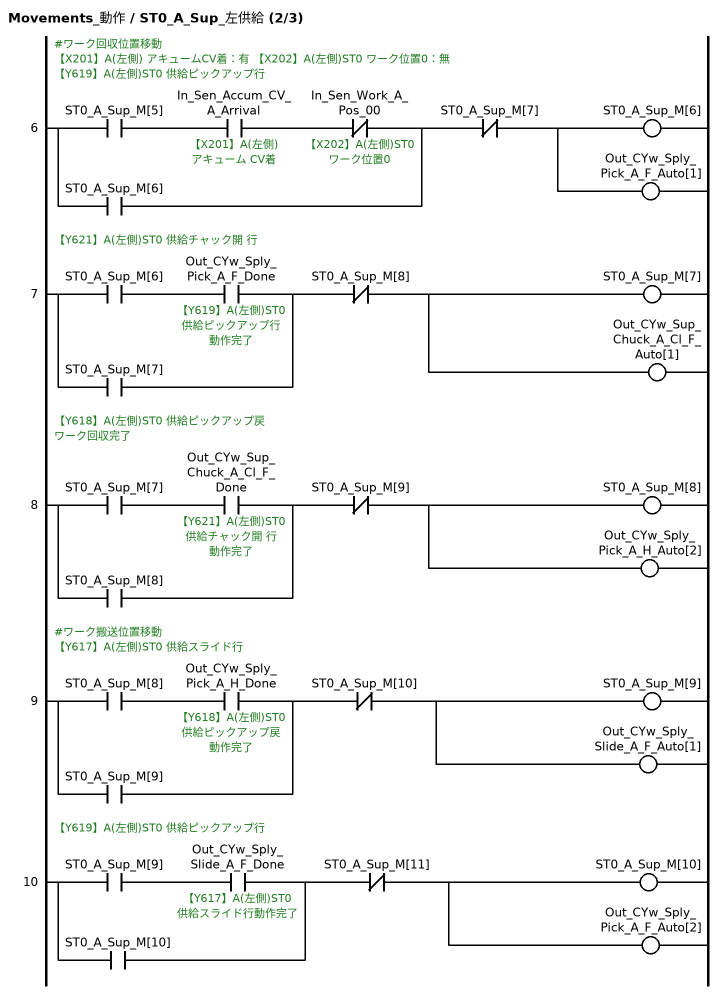
(* [picture p24: Movements_動作 / ST0_A_Sup_左供給, rungs 6-10] *)
(* Rung 6: #ワーク回収位置移動 / 【X201】A(左側) アキュームCV着：有 【X202】A(左側)ST0 ワーク位置0：無 / 【Y619】A(左側)ST0 供給ピックアップ行 *)
_p20 := ((ST0_A_Sup_M[5] AND In_Sen_Accum_CV_A_Arrival AND NOT In_Sen_Work_A_Pos_00) OR ST0_A_Sup_M[6]) AND NOT ST0_A_Sup_M[7];
ST0_A_Sup_M[6] := _p20;
Out_CYw_Sply_Pick_A_F_Auto[1] := _p20;
(* Rung 7: 【Y621】A(左側)ST0 供給チャック開 行 *)
_p21 := ((ST0_A_Sup_M[6] AND Out_CYw_Sply_Pick_A_F_Done) OR ST0_A_Sup_M[7]) AND NOT ST0_A_Sup_M[8];
ST0_A_Sup_M[7] := _p21;
Out_CYw_Sup_Chuck_A_Cl_F_Auto[1] := _p21;
(* Rung 8: 【Y618】A(左側)ST0 供給ピックアップ戻 / ワーク回収完了 *)
_p22 := ((ST0_A_Sup_M[7] AND Out_CYw_Sup_Chuck_A_Cl_F_Done) OR ST0_A_Sup_M[8]) AND NOT ST0_A_Sup_M[9];
ST0_A_Sup_M[8] := _p22;
Out_CYw_Sply_Pick_A_H_Auto[2] := _p22;
(* Rung 9: #ワーク搬送位置移動 / 【Y617】A(左側)ST0 供給スライド行 *)
_p23 := ((ST0_A_Sup_M[8] AND Out_CYw_Sply_Pick_A_H_Done) OR ST0_A_Sup_M[9]) AND NOT ST0_A_Sup_M[10];
ST0_A_Sup_M[9] := _p23;
Out_CYw_Sply_Slide_A_F_Auto[1] := _p23;
(* Rung 10: 【Y619】A(左側)ST0 供給ピックアップ行 *)
_p24 := ((ST0_A_Sup_M[9] AND Out_CYw_Sply_Slide_A_F_Done) OR ST0_A_Sup_M[10]) AND NOT ST0_A_Sup_M[11];
ST0_A_Sup_M[10] := _p24;
Out_CYw_Sply_Pick_A_F_Auto[2] := _p24;

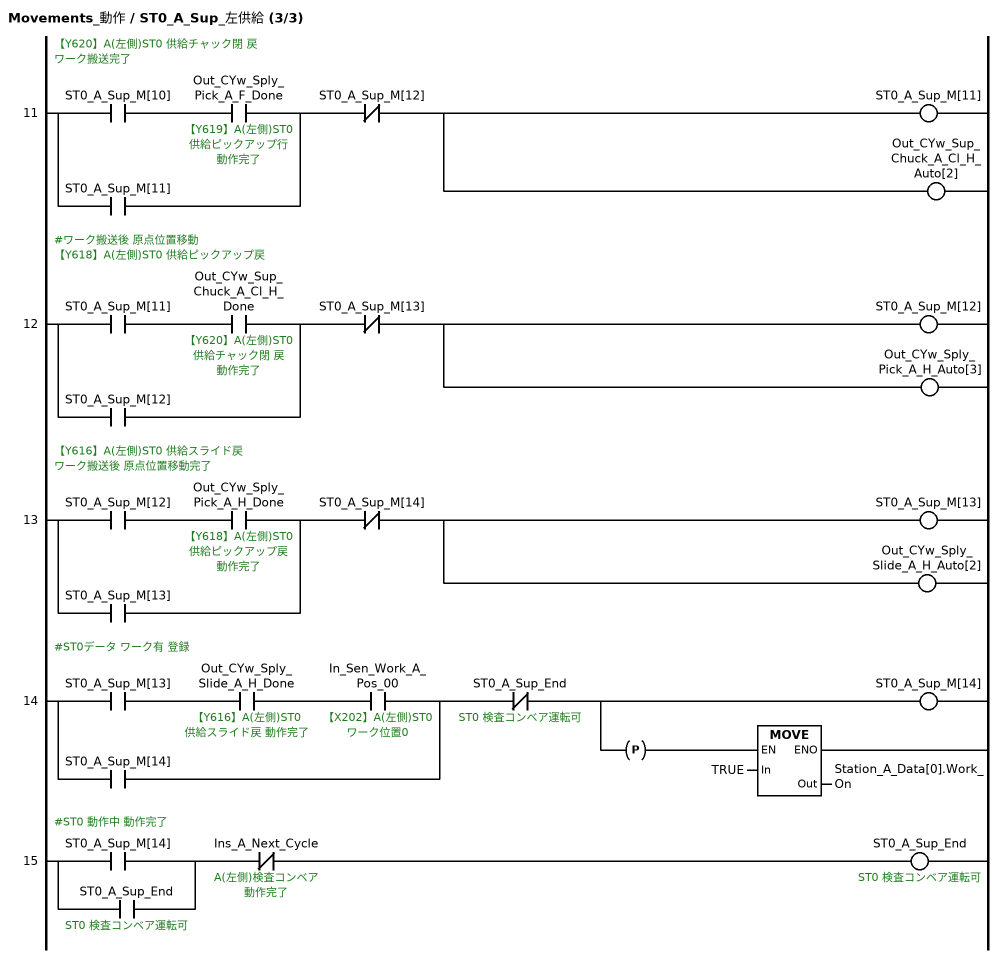
(* Rung 11: 【Y620】A(左側)ST0 供給チャック閉 戻 / ワーク搬送完了 *)
_p25 := ((ST0_A_Sup_M[10] AND Out_CYw_Sply_Pick_A_F_Done) OR ST0_A_Sup_M[11]) AND NOT ST0_A_Sup_M[12];
ST0_A_Sup_M[11] := _p25;
Out_CYw_Sup_Chuck_A_Cl_H_Auto[2] := _p25;
(* Rung 12: #ワーク搬送後 原点位置移動 / 【Y618】A(左側)ST0 供給ピックアップ戻 *)
_p26 := ((ST0_A_Sup_M[11] AND Out_CYw_Sup_Chuck_A_Cl_H_Done) OR ST0_A_Sup_M[12]) AND NOT ST0_A_Sup_M[13];
ST0_A_Sup_M[12] := _p26;
Out_CYw_Sply_Pick_A_H_Auto[3] := _p26;
(* Rung 13: 【Y616】A(左側)ST0 供給スライド戻 / ワーク搬送後 原点位置移動完了 *)
_p27 := ((ST0_A_Sup_M[12] AND Out_CYw_Sply_Pick_A_H_Done) OR ST0_A_Sup_M[13]) AND NOT ST0_A_Sup_M[14];
ST0_A_Sup_M[13] := _p27;
Out_CYw_Sply_Slide_A_H_Auto[2] := _p27;
(* Rung 14: #ST0データ ワーク有 登録 *)
_p28 := ((ST0_A_Sup_M[13] AND Out_CYw_Sply_Slide_A_H_Done AND In_Sen_Work_A_Pos_00) OR ST0_A_Sup_M[14]) AND NOT ST0_A_Sup_End;
ST0_A_Sup_M[14] := _p28;
_e29(CLK := _p28);
IF _e29.Q THEN Station_A_Data[0].Work_On := TRUE; END_IF;
(* Rung 15: #ST0 動作中 動作完了 *)
ST0_A_Sup_End := (ST0_A_Sup_M[14] OR ST0_A_Sup_End) AND NOT Ins_A_Next_Cycle;

(* Section ST1_A_Ca1_左Ca1検査: ladder, written here as Structured Text *)

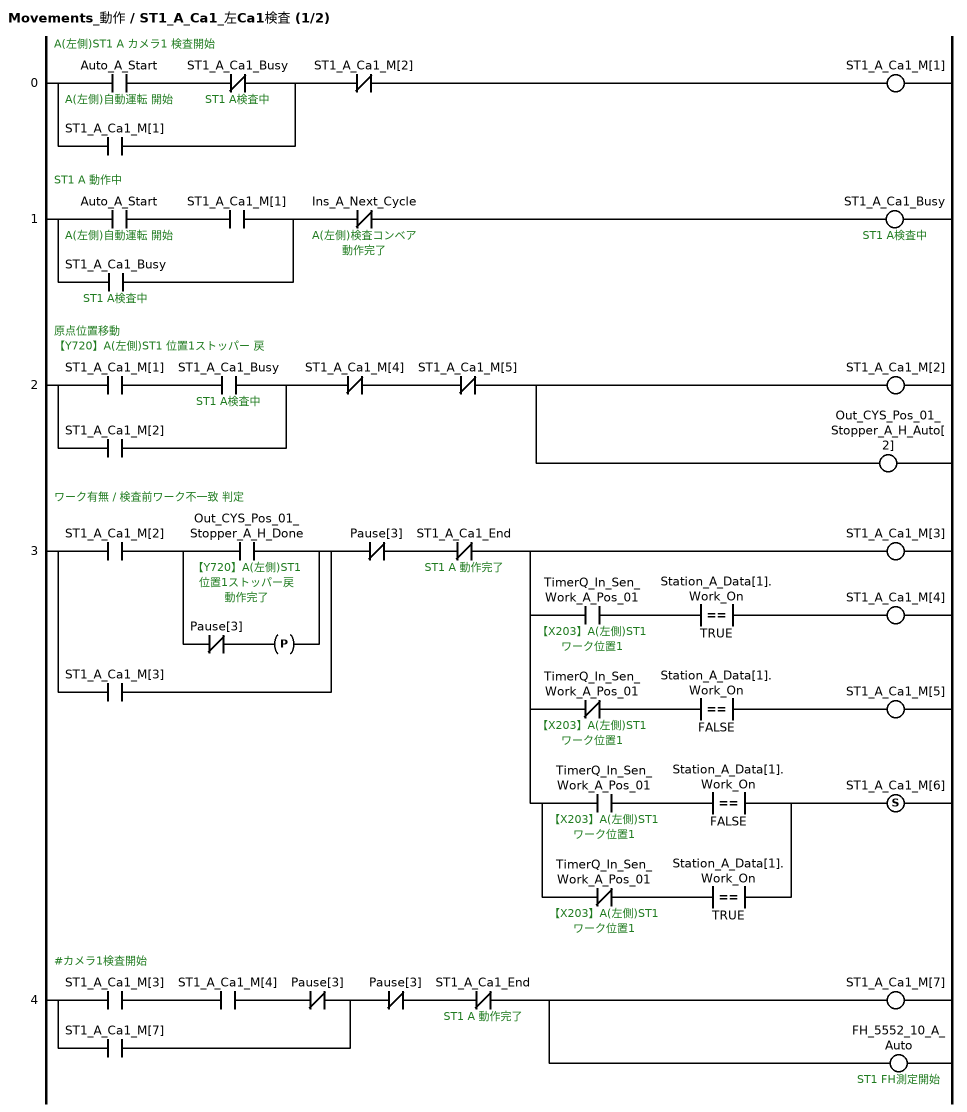
(* Rung 0: A(左側)ST1 A カメラ1 検査開始 *)
ST1_A_Ca1_M[1] := ((Auto_A_Start AND NOT ST1_A_Ca1_Busy) OR ST1_A_Ca1_M[1]) AND NOT ST1_A_Ca1_M[2];
(* Rung 1: ST1 A 動作中 *)
ST1_A_Ca1_Busy := ((Auto_A_Start AND ST1_A_Ca1_M[1]) OR ST1_A_Ca1_Busy) AND NOT Ins_A_Next_Cycle;
(* Rung 2: 原点位置移動 / 【Y720】A(左側)ST1 位置1ストッパー 戻 *)
_p30 := ((ST1_A_Ca1_M[1] AND ST1_A_Ca1_Busy) OR ST1_A_Ca1_M[2]) AND NOT ST1_A_Ca1_M[4] AND NOT ST1_A_Ca1_M[5];
ST1_A_Ca1_M[2] := _p30;
Out_CYS_Pos_01_Stopper_A_H_Auto[2] := _p30;
(* Rung 3: ワーク有無 / 検査前ワーク不一致 判定 *)
_e31(CLK := ST1_A_Ca1_M[2] AND NOT Pause[3]);
_p32 := ((ST1_A_Ca1_M[2] AND Out_CYS_Pos_01_Stopper_A_H_Done) OR _e31.Q OR ST1_A_Ca1_M[3]) AND NOT Pause[3] AND NOT ST1_A_Ca1_End;
ST1_A_Ca1_M[3] := _p32;
ST1_A_Ca1_M[4] := _p32 AND TimerQ_In_Sen_Work_A_Pos_01 AND (Station_A_Data[1].Work_On = TRUE);
ST1_A_Ca1_M[5] := _p32 AND NOT TimerQ_In_Sen_Work_A_Pos_01 AND (Station_A_Data[1].Work_On = FALSE);
IF _p32 AND ((TimerQ_In_Sen_Work_A_Pos_01 AND (Station_A_Data[1].Work_On = FALSE)) OR (NOT TimerQ_In_Sen_Work_A_Pos_01 AND (Station_A_Data[1].Work_On = TRUE))) THEN
    ST1_A_Ca1_M[6] := TRUE;
END_IF;
(* Rung 4: #カメラ1検査開始 *)
_p33 := ((ST1_A_Ca1_M[3] AND ST1_A_Ca1_M[4] AND NOT Pause[3]) OR ST1_A_Ca1_M[7]) AND NOT Pause[3] AND NOT ST1_A_Ca1_End;
ST1_A_Ca1_M[7] := _p33;
FH_5552_10_A_Auto := _p33;

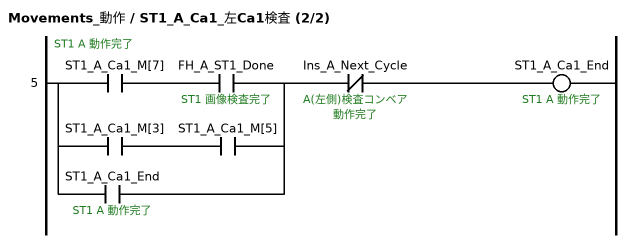
(* Rung 5: ST1 A 動作完了 *)
ST1_A_Ca1_End := ((ST1_A_Ca1_M[7] AND FH_A_ST1_Done) OR (ST1_A_Ca1_M[3] AND ST1_A_Ca1_M[5]) OR ST1_A_Ca1_End) AND NOT Ins_A_Next_Cycle;

(* Section ST2_A_Hgt_左高さ検査: ladder, written here as Structured Text *)

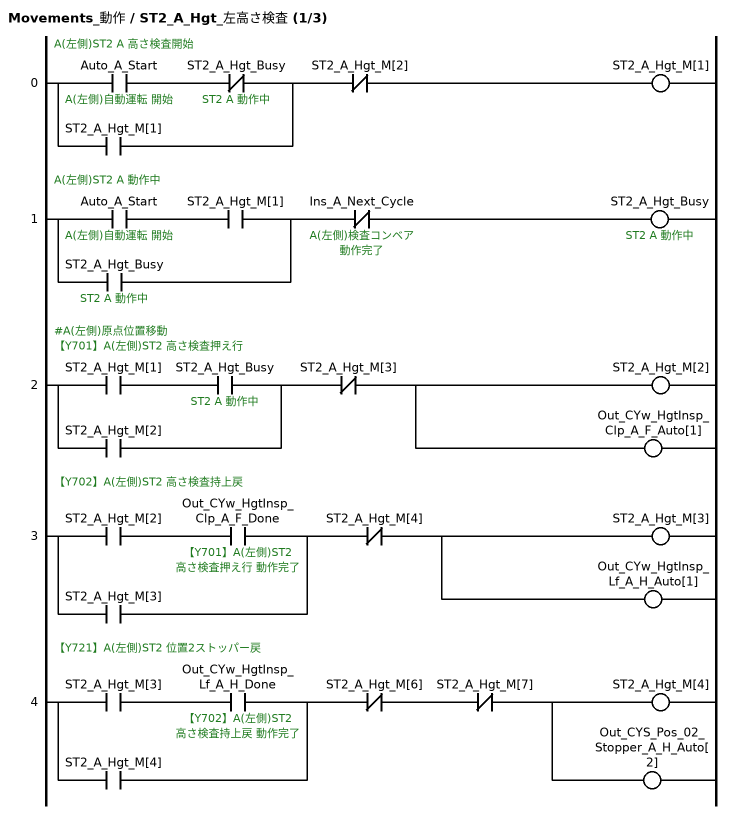
(* Rung 0: A(左側)ST2 A 高さ検査開始 *)
ST2_A_Hgt_M[1] := ((Auto_A_Start AND NOT ST2_A_Hgt_Busy) OR ST2_A_Hgt_M[1]) AND NOT ST2_A_Hgt_M[2];
(* Rung 1: A(左側)ST2 A 動作中 *)
ST2_A_Hgt_Busy := ((Auto_A_Start AND ST2_A_Hgt_M[1]) OR ST2_A_Hgt_Busy) AND NOT Ins_A_Next_Cycle;
(* Rung 2: #A(左側)原点位置移動 / 【Y701】A(左側)ST2 高さ検査押え行 *)
_p34 := ((ST2_A_Hgt_M[1] AND ST2_A_Hgt_Busy) OR ST2_A_Hgt_M[2]) AND NOT ST2_A_Hgt_M[3];
ST2_A_Hgt_M[2] := _p34;
Out_CYw_HgtInsp_Clp_A_F_Auto[1] := _p34;
(* Rung 3: 【Y702】A(左側)ST2 高さ検査持上戻 *)
_p35 := ((ST2_A_Hgt_M[2] AND Out_CYw_HgtInsp_Clp_A_F_Done) OR ST2_A_Hgt_M[3]) AND NOT ST2_A_Hgt_M[4];
ST2_A_Hgt_M[3] := _p35;
Out_CYw_HgtInsp_Lf_A_H_Auto[1] := _p35;
(* Rung 4: 【Y721】A(左側)ST2 位置2ストッパー戻 *)
_p36 := ((ST2_A_Hgt_M[3] AND Out_CYw_HgtInsp_Lf_A_H_Done) OR ST2_A_Hgt_M[4]) AND NOT ST2_A_Hgt_M[6] AND NOT ST2_A_Hgt_M[7];
ST2_A_Hgt_M[4] := _p36;
Out_CYS_Pos_02_Stopper_A_H_Auto[2] := _p36;

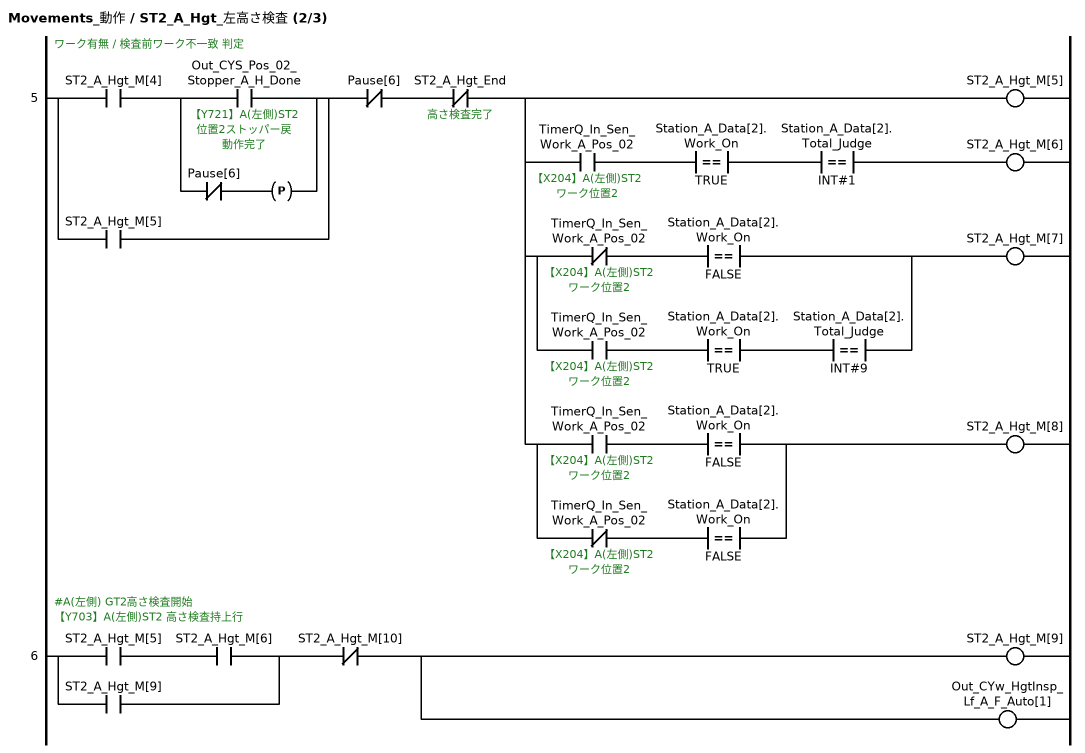
(* Rung 5: ワーク有無 / 検査前ワーク不一致 判定 *)
_e37(CLK := ST2_A_Hgt_M[4] AND NOT Pause[6]);
_p38 := ((ST2_A_Hgt_M[4] AND Out_CYS_Pos_02_Stopper_A_H_Done) OR _e37.Q OR ST2_A_Hgt_M[5]) AND NOT Pause[6] AND NOT ST2_A_Hgt_End;
ST2_A_Hgt_M[5] := _p38;
ST2_A_Hgt_M[6] := _p38 AND TimerQ_In_Sen_Work_A_Pos_02 AND (Station_A_Data[2].Work_On = TRUE) AND (Station_A_Data[2].Total_Judge = INT#1);
ST2_A_Hgt_M[7] := _p38 AND ((NOT TimerQ_In_Sen_Work_A_Pos_02 AND (Station_A_Data[2].Work_On = FALSE)) OR (TimerQ_In_Sen_Work_A_Pos_02 AND (Station_A_Data[2].Work_On = TRUE) AND (Station_A_Data[2].Total_Judge = INT#9)));
ST2_A_Hgt_M[8] := _p38 AND ((TimerQ_In_Sen_Work_A_Pos_02 AND (Station_A_Data[2].Work_On = FALSE)) OR (NOT TimerQ_In_Sen_Work_A_Pos_02 AND (Station_A_Data[2].Work_On = FALSE)));
(* Rung 6: #A(左側) GT2高さ検査開始 / 【Y703】A(左側)ST2 高さ検査持上行 *)
_p39 := ((ST2_A_Hgt_M[5] AND ST2_A_Hgt_M[6]) OR ST2_A_Hgt_M[9]) AND NOT ST2_A_Hgt_M[10];
ST2_A_Hgt_M[9] := _p39;
Out_CYw_HgtInsp_Lf_A_F_Auto[1] := _p39;

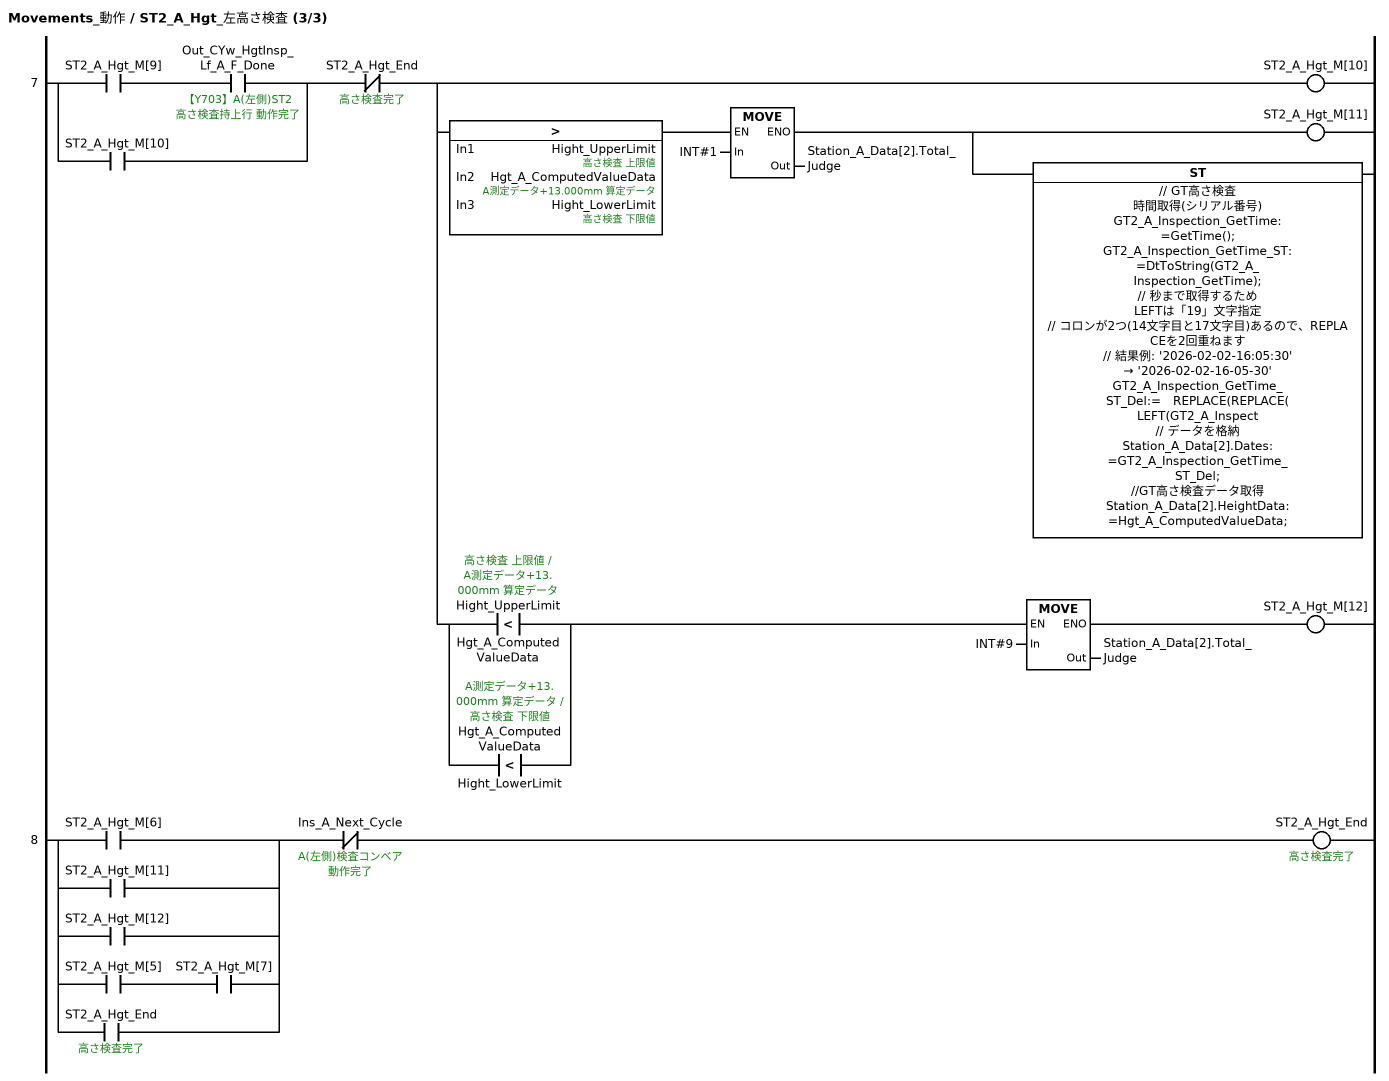
(* Rung 7 *)
_p40 := ((ST2_A_Hgt_M[9] AND Out_CYw_HgtInsp_Lf_A_F_Done) OR ST2_A_Hgt_M[10]) AND NOT ST2_A_Hgt_End;
ST2_A_Hgt_M[10] := _p40;
IF _p40 AND GT(Hight_UpperLimit, Hgt_A_ComputedValueData, Hight_LowerLimit) THEN
    Station_A_Data[2].Total_Judge := INT#1;
END_IF;
_p41 := _p40 AND GT(Hight_UpperLimit, Hgt_A_ComputedValueData, Hight_LowerLimit);
ST2_A_Hgt_M[11] := _p41;
IF _p41 THEN
    // GT高さ検査 時間取得(シリアル番号)
    GT2_A_Inspection_GetTime:=GetTime();
    GT2_A_Inspection_GetTime_ST:=DtToString(GT2_A_Inspection_GetTime);
    // 秒まで取得するため LEFTは「19」文字指定
    // コロンが2つ(14文字目と17文字目)あるので、REPLACEを2回重ねます
    // 結果例: '2026-02-02-16:05:30' → '2026-02-02-16-05-30'
    GT2_A_Inspection_GetTime_ST_Del:=   REPLACE(REPLACE(LEFT(GT2_A_Inspection_GetTime_ST, UINT#19), STRING#'-', UINT#1, UINT#17), STRING#'-', UINT#1, UINT#14);
    // データを格納
    Station_A_Data[2].Dates:=GT2_A_Inspection_GetTime_ST_Del;
    //GT高さ検査データ取得
    Station_A_Data[2].HeightData:=Hgt_A_ComputedValueData;
END_IF;
IF _p40 AND ((Hight_UpperLimit < Hgt_A_ComputedValueData) OR (Hgt_A_ComputedValueData < Hight_LowerLimit)) THEN
    Station_A_Data[2].Total_Judge := INT#9;
END_IF;
ST2_A_Hgt_M[12] := _p40 AND ((Hight_UpperLimit < Hgt_A_ComputedValueData) OR (Hgt_A_ComputedValueData < Hight_LowerLimit));
(* Rung 8 *)
ST2_A_Hgt_End := (ST2_A_Hgt_M[6] OR ST2_A_Hgt_M[11] OR ST2_A_Hgt_M[12] OR (ST2_A_Hgt_M[5] AND ST2_A_Hgt_M[7]) OR ST2_A_Hgt_End) AND NOT Ins_A_Next_Cycle;

(* Section ST3_A_Dis1_左NG1排出: ladder, written here as Structured Text *)

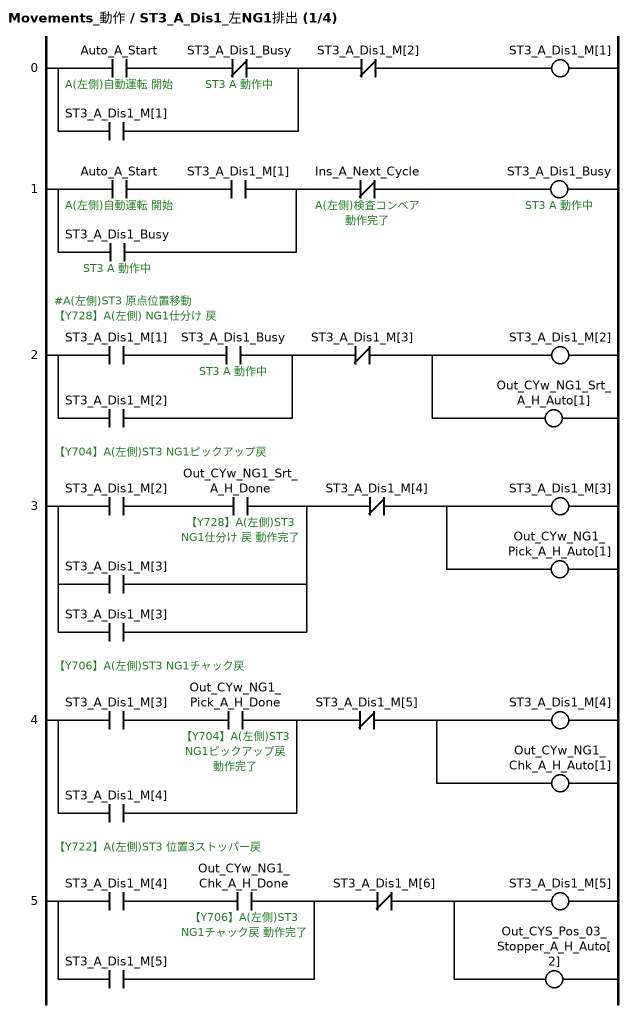
(* Rung 0 *)
ST3_A_Dis1_M[1] := ((Auto_A_Start AND NOT ST3_A_Dis1_Busy) OR ST3_A_Dis1_M[1]) AND NOT ST3_A_Dis1_M[2];
(* Rung 1 *)
ST3_A_Dis1_Busy := ((Auto_A_Start AND ST3_A_Dis1_M[1]) OR ST3_A_Dis1_Busy) AND NOT Ins_A_Next_Cycle;
(* Rung 2: #A(左側)ST3 原点位置移動 / 【Y728】A(左側) NG1仕分け 戻 *)
_p42 := ((ST3_A_Dis1_M[1] AND ST3_A_Dis1_Busy) OR ST3_A_Dis1_M[2]) AND NOT ST3_A_Dis1_M[3];
ST3_A_Dis1_M[2] := _p42;
Out_CYw_NG1_Srt_A_H_Auto[1] := _p42;
(* Rung 3: 【Y704】A(左側)ST3 NG1ピックアップ戻 *)
_p43 := ((ST3_A_Dis1_M[2] AND Out_CYw_NG1_Srt_A_H_Done) OR ST3_A_Dis1_M[3] OR ST3_A_Dis1_M[3]) AND NOT ST3_A_Dis1_M[4];
ST3_A_Dis1_M[3] := _p43;
Out_CYw_NG1_Pick_A_H_Auto[1] := _p43;
(* Rung 4: 【Y706】A(左側)ST3 NG1チャック戻 *)
_p44 := ((ST3_A_Dis1_M[3] AND Out_CYw_NG1_Pick_A_H_Done) OR ST3_A_Dis1_M[4]) AND NOT ST3_A_Dis1_M[5];
ST3_A_Dis1_M[4] := _p44;
Out_CYw_NG1_Chk_A_H_Auto[1] := _p44;
(* Rung 5: 【Y722】A(左側)ST3 位置3ストッパー戻 *)
_p45 := ((ST3_A_Dis1_M[4] AND Out_CYw_NG1_Chk_A_H_Done) OR ST3_A_Dis1_M[5]) AND NOT ST3_A_Dis1_M[6];
ST3_A_Dis1_M[5] := _p45;
Out_CYS_Pos_03_Stopper_A_H_Auto[2] := _p45;

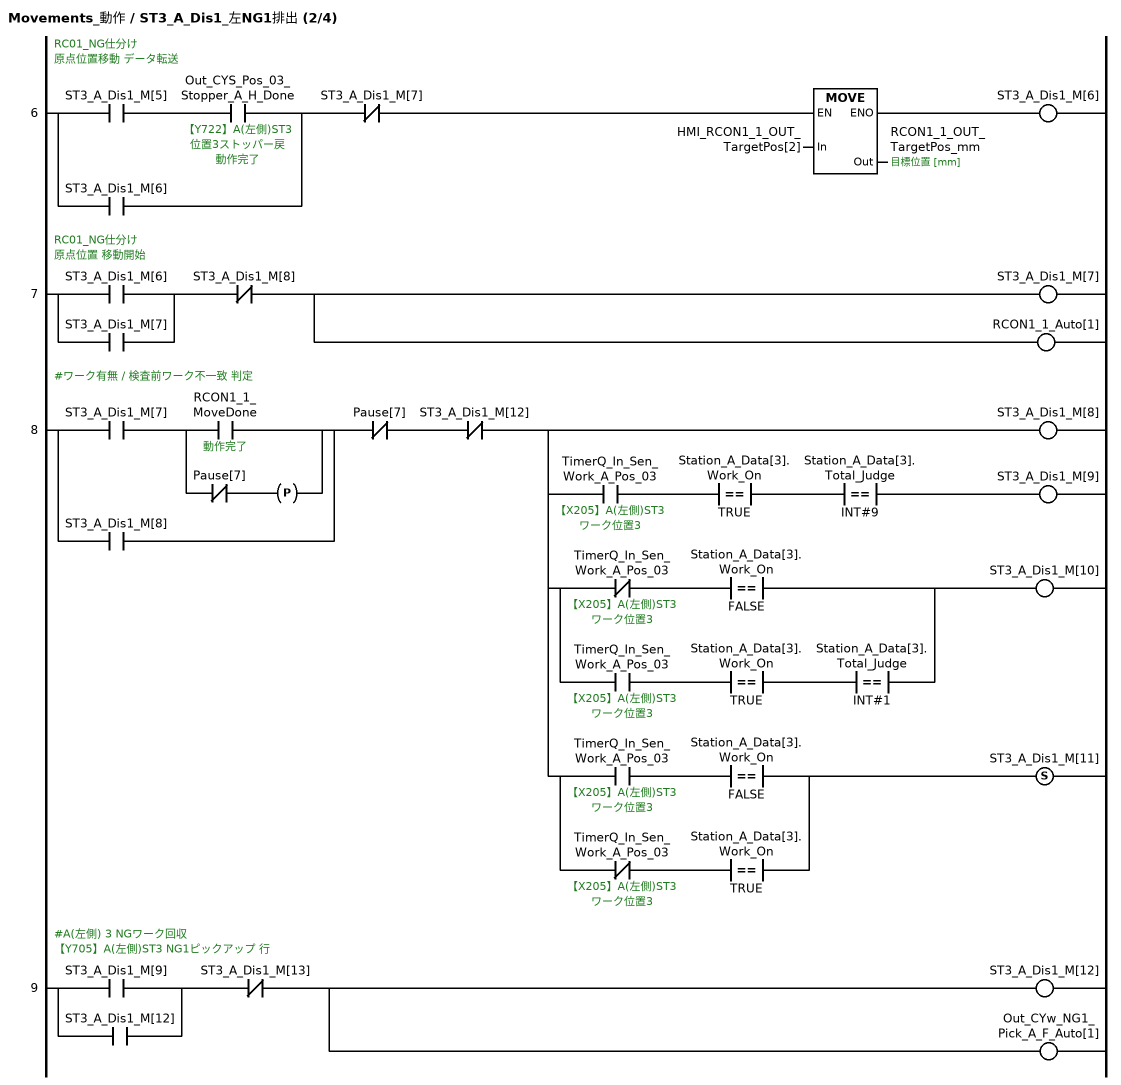
(* Rung 6: RC01_NG仕分け / 原点位置移動 データ転送 *)
IF ((ST3_A_Dis1_M[5] AND Out_CYS_Pos_03_Stopper_A_H_Done) OR ST3_A_Dis1_M[6]) AND NOT ST3_A_Dis1_M[7] THEN
    RCON1_1_OUT_TargetPos_mm := HMI_RCON1_1_OUT_TargetPos[2];
END_IF;
ST3_A_Dis1_M[6] := ((ST3_A_Dis1_M[5] AND Out_CYS_Pos_03_Stopper_A_H_Done) OR ST3_A_Dis1_M[6]) AND NOT ST3_A_Dis1_M[7];
(* Rung 7: RC01_NG仕分け / 原点位置 移動開始 *)
_p46 := (ST3_A_Dis1_M[6] OR ST3_A_Dis1_M[7]) AND NOT ST3_A_Dis1_M[8];
ST3_A_Dis1_M[7] := _p46;
RCON1_1_Auto[1] := _p46;
(* Rung 8: #ワーク有無 / 検査前ワーク不一致 判定 *)
_e47(CLK := ST3_A_Dis1_M[7] AND NOT Pause[7]);
_p48 := ((ST3_A_Dis1_M[7] AND RCON1_1_MoveDone) OR _e47.Q OR ST3_A_Dis1_M[8]) AND NOT Pause[7] AND NOT ST3_A_Dis1_M[12];
ST3_A_Dis1_M[8] := _p48;
ST3_A_Dis1_M[9] := _p48 AND TimerQ_In_Sen_Work_A_Pos_03 AND (Station_A_Data[3].Work_On = TRUE) AND (Station_A_Data[3].Total_Judge = INT#9);
ST3_A_Dis1_M[10] := _p48 AND ((NOT TimerQ_In_Sen_Work_A_Pos_03 AND (Station_A_Data[3].Work_On = FALSE)) OR (TimerQ_In_Sen_Work_A_Pos_03 AND (Station_A_Data[3].Work_On = TRUE) AND (Station_A_Data[3].Total_Judge = INT#1)));
IF _p48 AND ((TimerQ_In_Sen_Work_A_Pos_03 AND (Station_A_Data[3].Work_On = FALSE)) OR (NOT TimerQ_In_Sen_Work_A_Pos_03 AND (Station_A_Data[3].Work_On = TRUE))) THEN
    ST3_A_Dis1_M[11] := TRUE;
END_IF;
(* Rung 9: #A(左側) 3 NGワーク回収 / 【Y705】A(左側)ST3 NG1ピックアップ 行 *)
_p49 := (ST3_A_Dis1_M[9] OR ST3_A_Dis1_M[12]) AND NOT ST3_A_Dis1_M[13];
ST3_A_Dis1_M[12] := _p49;
Out_CYw_NG1_Pick_A_F_Auto[1] := _p49;

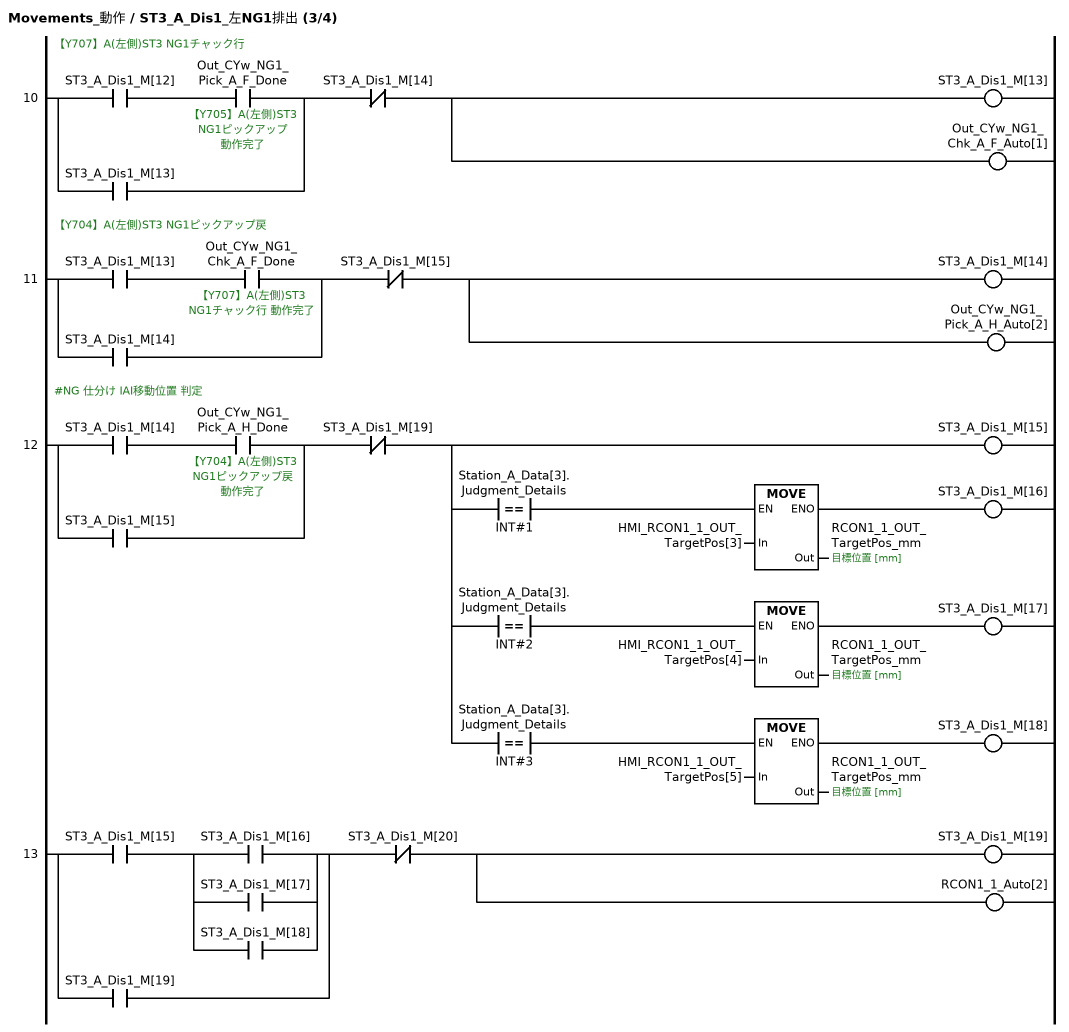
(* Rung 10: 【Y707】A(左側)ST3 NG1チャック行 *)
_p50 := ((ST3_A_Dis1_M[12] AND Out_CYw_NG1_Pick_A_F_Done) OR ST3_A_Dis1_M[13]) AND NOT ST3_A_Dis1_M[14];
ST3_A_Dis1_M[13] := _p50;
Out_CYw_NG1_Chk_A_F_Auto[1] := _p50;
(* Rung 11: 【Y704】A(左側)ST3 NG1ピックアップ戻 *)
_p51 := ((ST3_A_Dis1_M[13] AND Out_CYw_NG1_Chk_A_F_Done) OR ST3_A_Dis1_M[14]) AND NOT ST3_A_Dis1_M[15];
ST3_A_Dis1_M[14] := _p51;
Out_CYw_NG1_Pick_A_H_Auto[2] := _p51;
(* Rung 12: #NG 仕分け IAI移動位置 判定 *)
_p52 := ((ST3_A_Dis1_M[14] AND Out_CYw_NG1_Pick_A_H_Done) OR ST3_A_Dis1_M[15]) AND NOT ST3_A_Dis1_M[19];
ST3_A_Dis1_M[15] := _p52;
IF _p52 AND (Station_A_Data[3].Judgment_Details = INT#1) THEN
    RCON1_1_OUT_TargetPos_mm := HMI_RCON1_1_OUT_TargetPos[3];
END_IF;
ST3_A_Dis1_M[16] := _p52 AND (Station_A_Data[3].Judgment_Details = INT#1);
IF _p52 AND (Station_A_Data[3].Judgment_Details = INT#2) THEN
    RCON1_1_OUT_TargetPos_mm := HMI_RCON1_1_OUT_TargetPos[4];
END_IF;
ST3_A_Dis1_M[17] := _p52 AND (Station_A_Data[3].Judgment_Details = INT#2);
IF _p52 AND (Station_A_Data[3].Judgment_Details = INT#3) THEN
    RCON1_1_OUT_TargetPos_mm := HMI_RCON1_1_OUT_TargetPos[5];
END_IF;
ST3_A_Dis1_M[18] := _p52 AND (Station_A_Data[3].Judgment_Details = INT#3);
(* Rung 13 *)
_p53 := ((ST3_A_Dis1_M[15] AND (ST3_A_Dis1_M[16] OR ST3_A_Dis1_M[17] OR ST3_A_Dis1_M[18])) OR ST3_A_Dis1_M[19]) AND NOT ST3_A_Dis1_M[20];
ST3_A_Dis1_M[19] := _p53;
RCON1_1_Auto[2] := _p53;

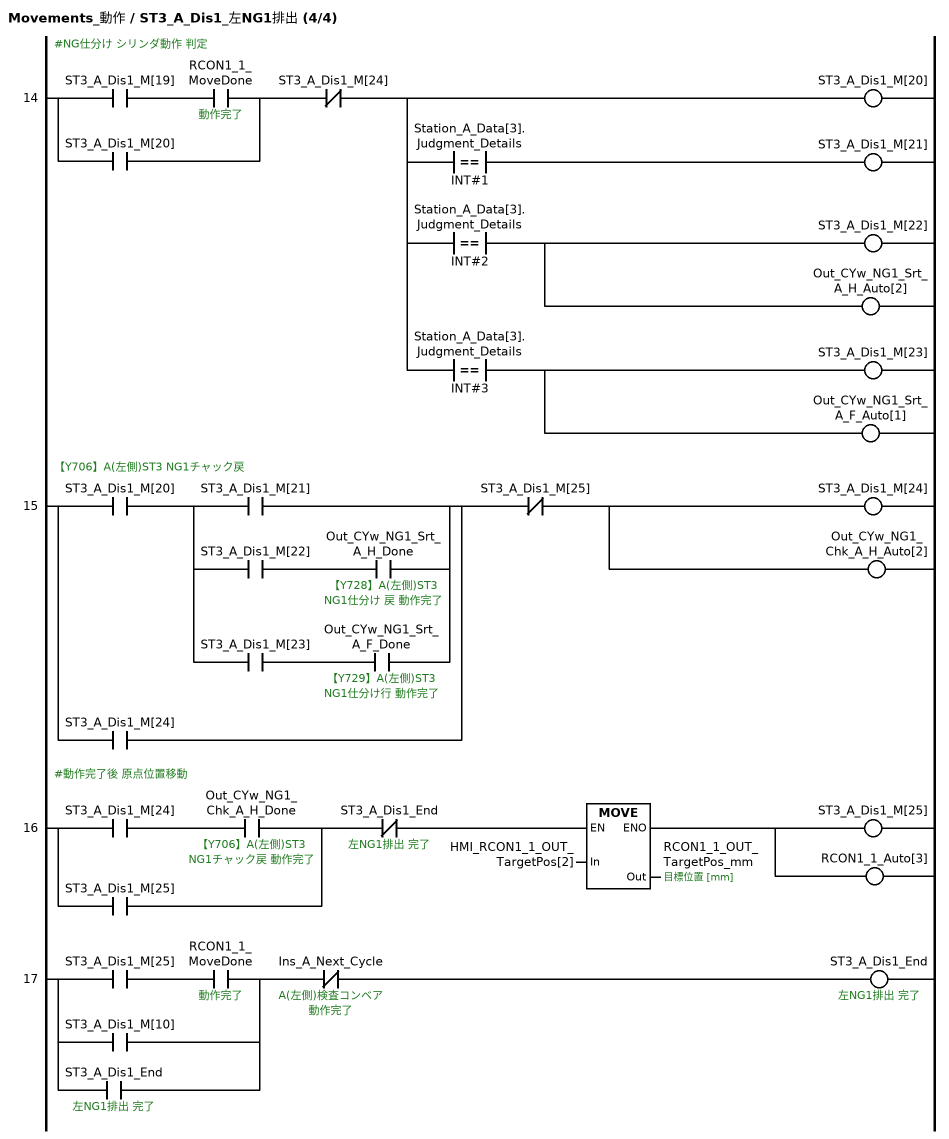
(* Rung 14: #NG仕分け シリンダ動作 判定 *)
_p54 := ((ST3_A_Dis1_M[19] AND RCON1_1_MoveDone) OR ST3_A_Dis1_M[20]) AND NOT ST3_A_Dis1_M[24];
ST3_A_Dis1_M[20] := _p54;
ST3_A_Dis1_M[21] := _p54 AND (Station_A_Data[3].Judgment_Details = INT#1);
_p55 := _p54 AND (Station_A_Data[3].Judgment_Details = INT#2);
ST3_A_Dis1_M[22] := _p55;
Out_CYw_NG1_Srt_A_H_Auto[2] := _p55;
_p56 := _p54 AND (Station_A_Data[3].Judgment_Details = INT#3);
ST3_A_Dis1_M[23] := _p56;
Out_CYw_NG1_Srt_A_F_Auto[1] := _p56;
(* Rung 15: 【Y706】A(左側)ST3 NG1チャック戻 *)
_p57 := ((ST3_A_Dis1_M[20] AND (ST3_A_Dis1_M[21] OR (ST3_A_Dis1_M[22] AND Out_CYw_NG1_Srt_A_H_Done) OR (ST3_A_Dis1_M[23] AND Out_CYw_NG1_Srt_A_F_Done))) OR ST3_A_Dis1_M[24]) AND NOT ST3_A_Dis1_M[25];
ST3_A_Dis1_M[24] := _p57;
Out_CYw_NG1_Chk_A_H_Auto[2] := _p57;
(* Rung 16: #動作完了後 原点位置移動 *)
IF ((ST3_A_Dis1_M[24] AND Out_CYw_NG1_Chk_A_H_Done) OR ST3_A_Dis1_M[25]) AND NOT ST3_A_Dis1_End THEN
    RCON1_1_OUT_TargetPos_mm := HMI_RCON1_1_OUT_TargetPos[2];
END_IF;
_p58 := ((ST3_A_Dis1_M[24] AND Out_CYw_NG1_Chk_A_H_Done) OR ST3_A_Dis1_M[25]) AND NOT ST3_A_Dis1_End;
ST3_A_Dis1_M[25] := _p58;
RCON1_1_Auto[3] := _p58;
(* Rung 17 *)
ST3_A_Dis1_End := ((ST3_A_Dis1_M[25] AND RCON1_1_MoveDone) OR ST3_A_Dis1_M[10] OR ST3_A_Dis1_End) AND NOT Ins_A_Next_Cycle;

(* Section ST4_A_Rev1_左反転1: ladder, written here as Structured Text *)

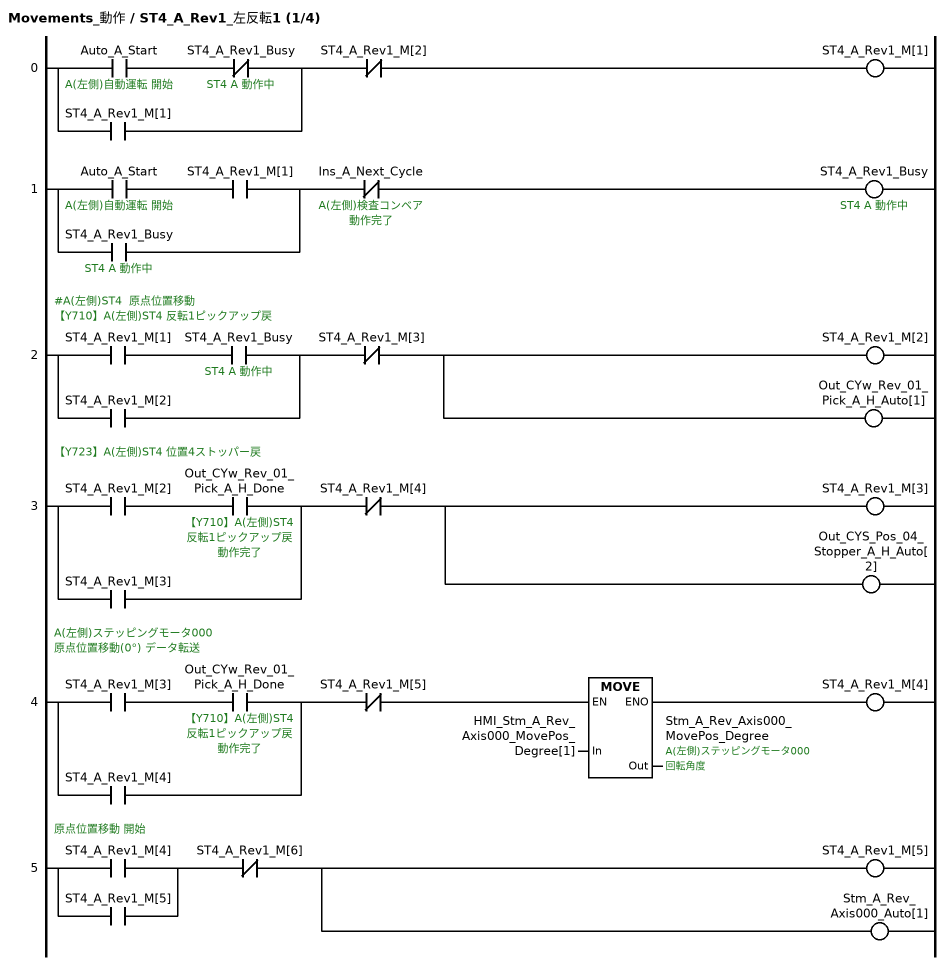
(* Rung 0 *)
ST4_A_Rev1_M[1] := ((Auto_A_Start AND NOT ST4_A_Rev1_Busy) OR ST4_A_Rev1_M[1]) AND NOT ST4_A_Rev1_M[2];
(* Rung 1 *)
ST4_A_Rev1_Busy := ((Auto_A_Start AND ST4_A_Rev1_M[1]) OR ST4_A_Rev1_Busy) AND NOT Ins_A_Next_Cycle;
(* Rung 2: #A(左側)ST4  原点位置移動 / 【Y710】A(左側)ST4 反転1ピックアップ戻 *)
_p59 := ((ST4_A_Rev1_M[1] AND ST4_A_Rev1_Busy) OR ST4_A_Rev1_M[2]) AND NOT ST4_A_Rev1_M[3];
ST4_A_Rev1_M[2] := _p59;
Out_CYw_Rev_01_Pick_A_H_Auto[1] := _p59;
(* Rung 3: 【Y723】A(左側)ST4 位置4ストッパー戻 *)
_p60 := ((ST4_A_Rev1_M[2] AND Out_CYw_Rev_01_Pick_A_H_Done) OR ST4_A_Rev1_M[3]) AND NOT ST4_A_Rev1_M[4];
ST4_A_Rev1_M[3] := _p60;
Out_CYS_Pos_04_Stopper_A_H_Auto[2] := _p60;
(* Rung 4: A(左側)ステッピングモータ000 / 原点位置移動(0°) データ転送 *)
IF ((ST4_A_Rev1_M[3] AND Out_CYw_Rev_01_Pick_A_H_Done) OR ST4_A_Rev1_M[4]) AND NOT ST4_A_Rev1_M[5] THEN
    Stm_A_Rev_Axis000_MovePos_Degree := HMI_Stm_A_Rev_Axis000_MovePos_Degree[1];
END_IF;
ST4_A_Rev1_M[4] := ((ST4_A_Rev1_M[3] AND Out_CYw_Rev_01_Pick_A_H_Done) OR ST4_A_Rev1_M[4]) AND NOT ST4_A_Rev1_M[5];
(* Rung 5: 原点位置移動 開始 *)
_p61 := (ST4_A_Rev1_M[4] OR ST4_A_Rev1_M[5]) AND NOT ST4_A_Rev1_M[6];
ST4_A_Rev1_M[5] := _p61;
Stm_A_Rev_Axis000_Auto[1] := _p61;

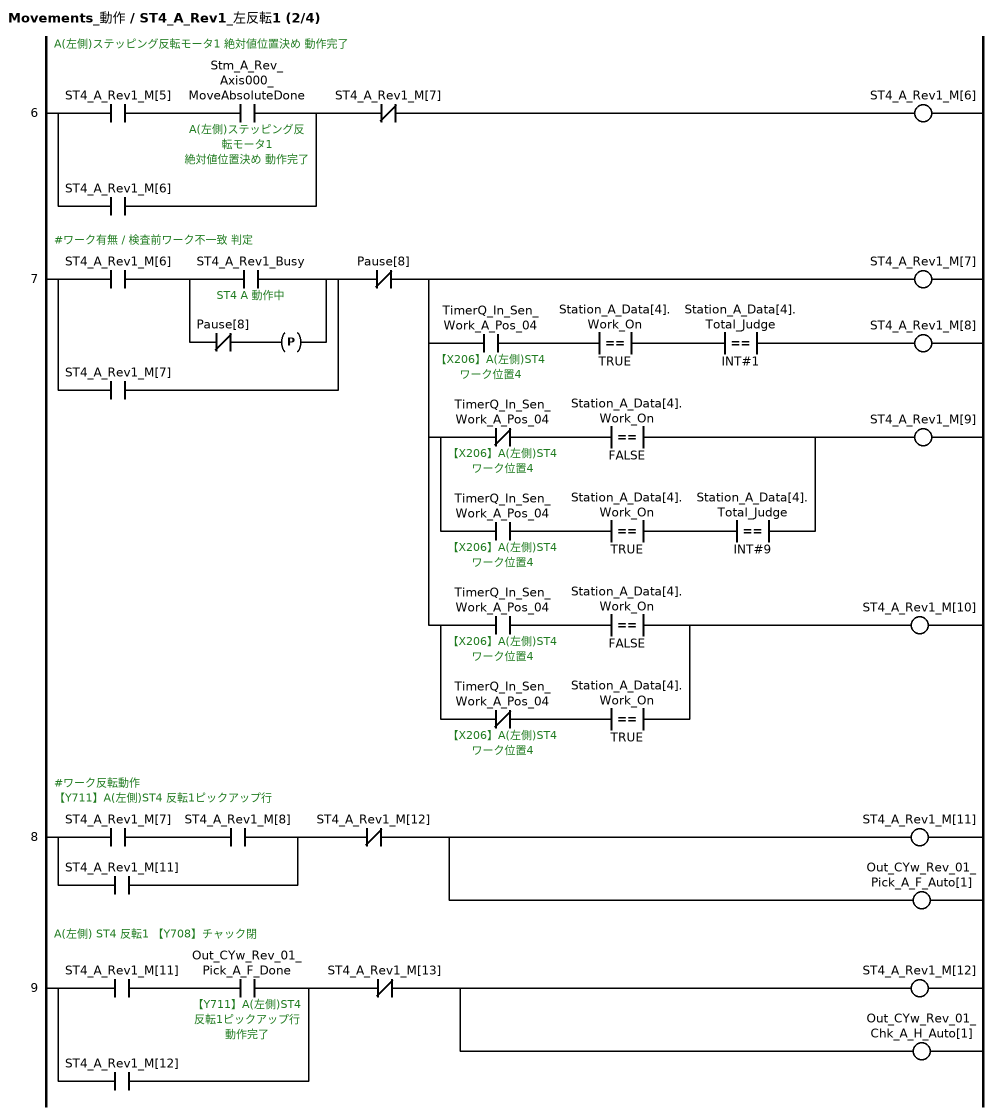
(* Rung 6: A(左側)ステッピング反転モータ1 絶対値位置決め 動作完了 *)
ST4_A_Rev1_M[6] := ((ST4_A_Rev1_M[5] AND Stm_A_Rev_Axis000_MoveAbsoluteDone) OR ST4_A_Rev1_M[6]) AND NOT ST4_A_Rev1_M[7];
(* Rung 7: #ワーク有無 / 検査前ワーク不一致 判定 *)
_e62(CLK := ST4_A_Rev1_M[6] AND NOT Pause[8]);
_p63 := ((ST4_A_Rev1_M[6] AND ST4_A_Rev1_Busy) OR _e62.Q OR ST4_A_Rev1_M[7]) AND NOT Pause[8];
ST4_A_Rev1_M[7] := _p63;
ST4_A_Rev1_M[8] := _p63 AND TimerQ_In_Sen_Work_A_Pos_04 AND (Station_A_Data[4].Work_On = TRUE) AND (Station_A_Data[4].Total_Judge = INT#1);
ST4_A_Rev1_M[9] := _p63 AND ((NOT TimerQ_In_Sen_Work_A_Pos_04 AND (Station_A_Data[4].Work_On = FALSE)) OR (TimerQ_In_Sen_Work_A_Pos_04 AND (Station_A_Data[4].Work_On = TRUE) AND (Station_A_Data[4].Total_Judge = INT#9)));
ST4_A_Rev1_M[10] := _p63 AND ((TimerQ_In_Sen_Work_A_Pos_04 AND (Station_A_Data[4].Work_On = FALSE)) OR (NOT TimerQ_In_Sen_Work_A_Pos_04 AND (Station_A_Data[4].Work_On = TRUE)));
(* Rung 8: #ワーク反転動作 / 【Y711】A(左側)ST4 反転1ピックアップ行 *)
_p64 := ((ST4_A_Rev1_M[7] AND ST4_A_Rev1_M[8]) OR ST4_A_Rev1_M[11]) AND NOT ST4_A_Rev1_M[12];
ST4_A_Rev1_M[11] := _p64;
Out_CYw_Rev_01_Pick_A_F_Auto[1] := _p64;
(* Rung 9: A(左側) ST4 反転1 【Y708】チャック閉 *)
_p65 := ((ST4_A_Rev1_M[11] AND Out_CYw_Rev_01_Pick_A_F_Done) OR ST4_A_Rev1_M[12]) AND NOT ST4_A_Rev1_M[13];
ST4_A_Rev1_M[12] := _p65;
Out_CYw_Rev_01_Chk_A_H_Auto[1] := _p65;

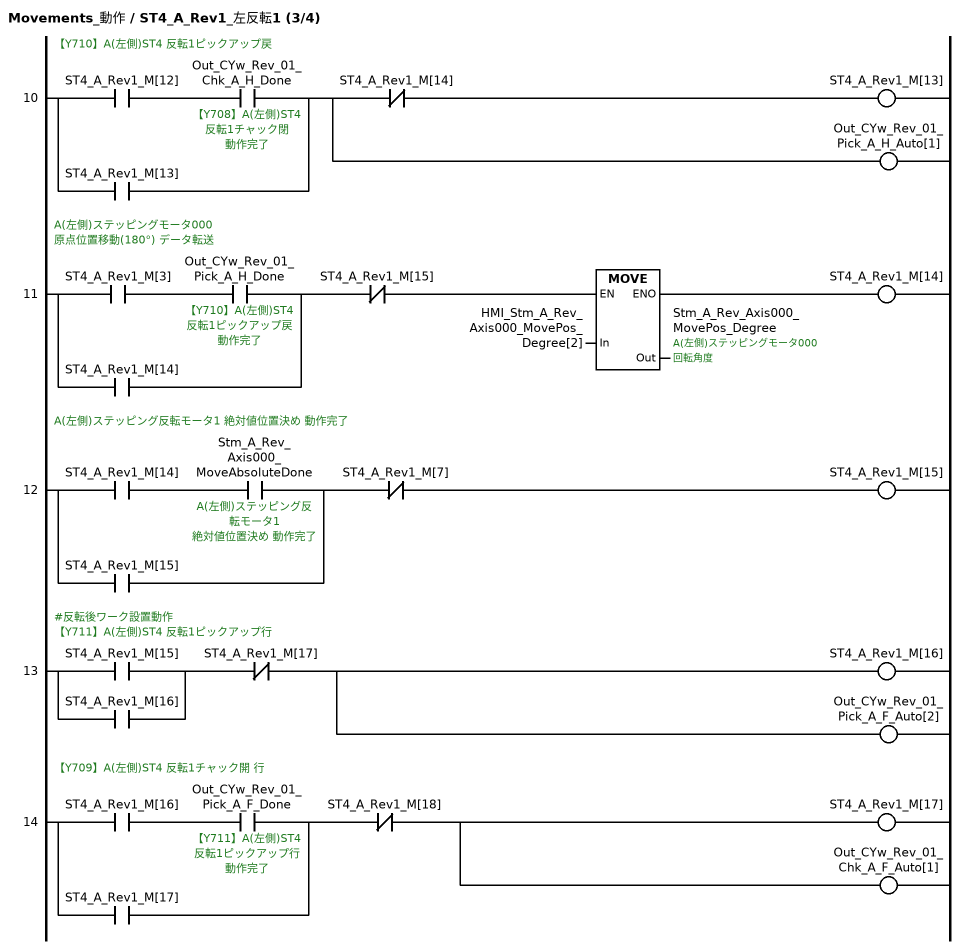
(* Rung 10: 【Y710】A(左側)ST4 反転1ピックアップ戻 *)
_p66 := (ST4_A_Rev1_M[12] AND Out_CYw_Rev_01_Chk_A_H_Done) OR ST4_A_Rev1_M[13];
ST4_A_Rev1_M[13] := _p66 AND NOT ST4_A_Rev1_M[14];
Out_CYw_Rev_01_Pick_A_H_Auto[1] := _p66;
(* Rung 11: A(左側)ステッピングモータ000 / 原点位置移動(180°) データ転送 *)
IF ((ST4_A_Rev1_M[3] AND Out_CYw_Rev_01_Pick_A_H_Done) OR ST4_A_Rev1_M[14]) AND NOT ST4_A_Rev1_M[15] THEN
    Stm_A_Rev_Axis000_MovePos_Degree := HMI_Stm_A_Rev_Axis000_MovePos_Degree[2];
END_IF;
ST4_A_Rev1_M[14] := ((ST4_A_Rev1_M[3] AND Out_CYw_Rev_01_Pick_A_H_Done) OR ST4_A_Rev1_M[14]) AND NOT ST4_A_Rev1_M[15];
(* Rung 12: A(左側)ステッピング反転モータ1 絶対値位置決め 動作完了 *)
ST4_A_Rev1_M[15] := ((ST4_A_Rev1_M[14] AND Stm_A_Rev_Axis000_MoveAbsoluteDone) OR ST4_A_Rev1_M[15]) AND NOT ST4_A_Rev1_M[7];
(* Rung 13: #反転後ワーク設置動作 / 【Y711】A(左側)ST4 反転1ピックアップ行 *)
_p67 := (ST4_A_Rev1_M[15] OR ST4_A_Rev1_M[16]) AND NOT ST4_A_Rev1_M[17];
ST4_A_Rev1_M[16] := _p67;
Out_CYw_Rev_01_Pick_A_F_Auto[2] := _p67;
(* Rung 14: 【Y709】A(左側)ST4 反転1チャック開 行 *)
_p68 := ((ST4_A_Rev1_M[16] AND Out_CYw_Rev_01_Pick_A_F_Done) OR ST4_A_Rev1_M[17]) AND NOT ST4_A_Rev1_M[18];
ST4_A_Rev1_M[17] := _p68;
Out_CYw_Rev_01_Chk_A_F_Auto[1] := _p68;

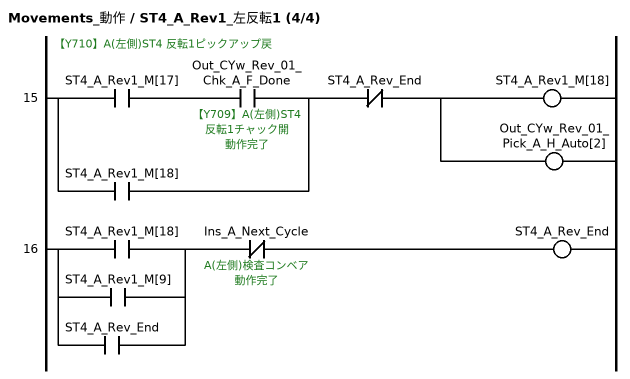
(* Rung 15: 【Y710】A(左側)ST4 反転1ピックアップ戻 *)
_p69 := ((ST4_A_Rev1_M[17] AND Out_CYw_Rev_01_Chk_A_F_Done) OR ST4_A_Rev1_M[18]) AND NOT ST4_A_Rev_End;
ST4_A_Rev1_M[18] := _p69;
Out_CYw_Rev_01_Pick_A_H_Auto[2] := _p69;
(* Rung 16 *)
ST4_A_Rev_End := (ST4_A_Rev1_M[18] OR ST4_A_Rev1_M[9] OR ST4_A_Rev_End) AND NOT Ins_A_Next_Cycle;

(* Section ST5_A_Ca2_左Ca2検査: ladder, written here as Structured Text *)

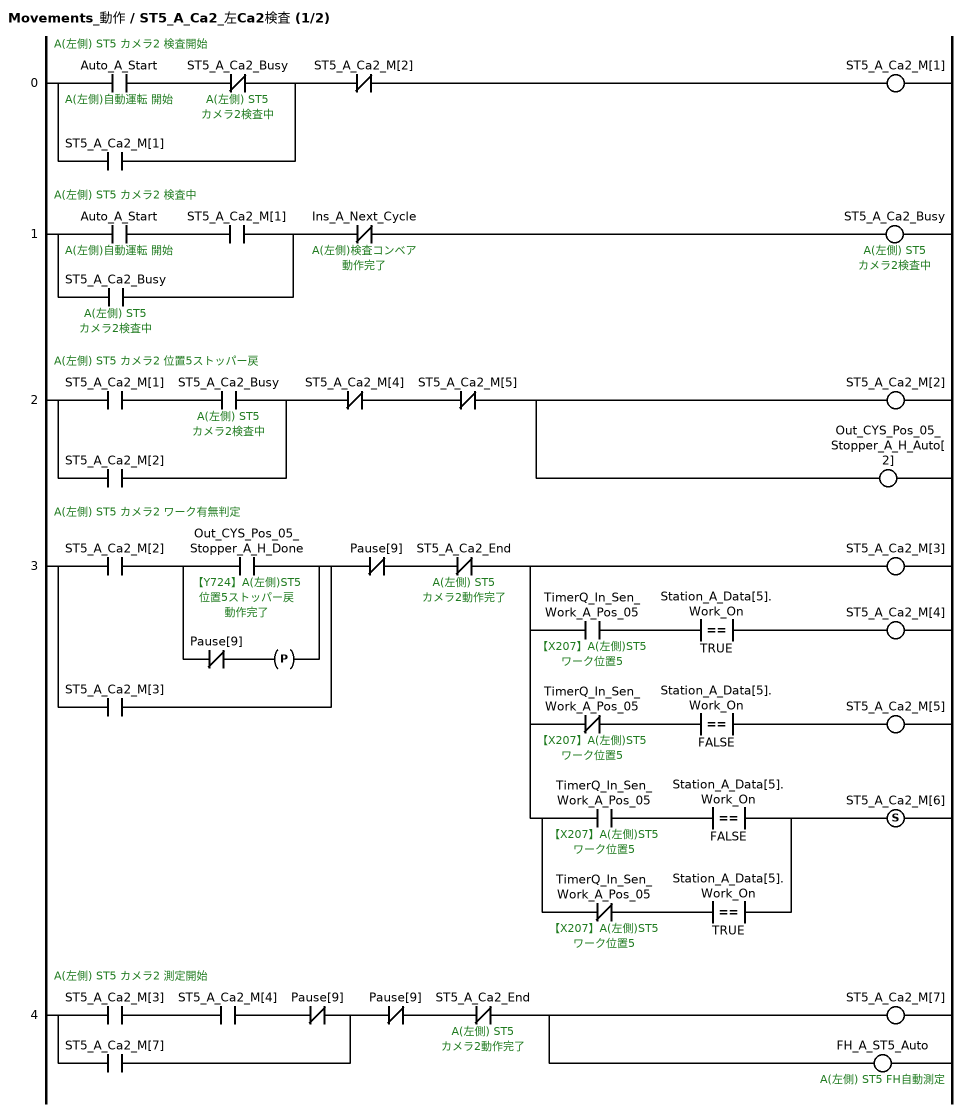
(* Rung 0: A(左側) ST5 カメラ2 検査開始 *)
ST5_A_Ca2_M[1] := ((Auto_A_Start AND NOT ST5_A_Ca2_Busy) OR ST5_A_Ca2_M[1]) AND NOT ST5_A_Ca2_M[2];
(* Rung 1: A(左側) ST5 カメラ2 検査中 *)
ST5_A_Ca2_Busy := ((Auto_A_Start AND ST5_A_Ca2_M[1]) OR ST5_A_Ca2_Busy) AND NOT Ins_A_Next_Cycle;
(* Rung 2: A(左側) ST5 カメラ2 位置5ストッパー戻 *)
_p70 := ((ST5_A_Ca2_M[1] AND ST5_A_Ca2_Busy) OR ST5_A_Ca2_M[2]) AND NOT ST5_A_Ca2_M[4] AND NOT ST5_A_Ca2_M[5];
ST5_A_Ca2_M[2] := _p70;
Out_CYS_Pos_05_Stopper_A_H_Auto[2] := _p70;
(* Rung 3: A(左側) ST5 カメラ2 ワーク有無判定 *)
_e71(CLK := ST5_A_Ca2_M[2] AND NOT Pause[9]);
_p72 := ((ST5_A_Ca2_M[2] AND Out_CYS_Pos_05_Stopper_A_H_Done) OR _e71.Q OR ST5_A_Ca2_M[3]) AND NOT Pause[9] AND NOT ST5_A_Ca2_End;
ST5_A_Ca2_M[3] := _p72;
ST5_A_Ca2_M[4] := _p72 AND TimerQ_In_Sen_Work_A_Pos_05 AND (Station_A_Data[5].Work_On = TRUE);
ST5_A_Ca2_M[5] := _p72 AND NOT TimerQ_In_Sen_Work_A_Pos_05 AND (Station_A_Data[5].Work_On = FALSE);
IF _p72 AND ((TimerQ_In_Sen_Work_A_Pos_05 AND (Station_A_Data[5].Work_On = FALSE)) OR (NOT TimerQ_In_Sen_Work_A_Pos_05 AND (Station_A_Data[5].Work_On = TRUE))) THEN
    ST5_A_Ca2_M[6] := TRUE;
END_IF;
(* Rung 4: A(左側) ST5 カメラ2 測定開始 *)
_p73 := ((ST5_A_Ca2_M[3] AND ST5_A_Ca2_M[4] AND NOT Pause[9]) OR ST5_A_Ca2_M[7]) AND NOT Pause[9] AND NOT ST5_A_Ca2_End;
ST5_A_Ca2_M[7] := _p73;
FH_A_ST5_Auto := _p73;

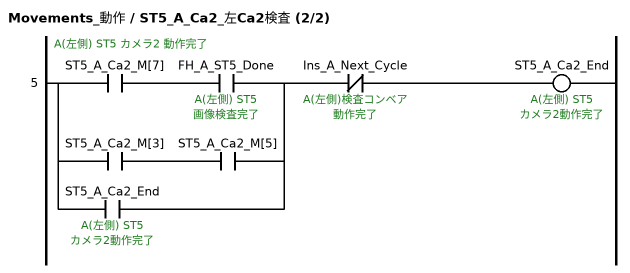
(* Rung 5: A(左側) ST5 カメラ2 動作完了 *)
ST5_A_Ca2_End := ((ST5_A_Ca2_M[7] AND FH_A_ST5_Done) OR (ST5_A_Ca2_M[3] AND ST5_A_Ca2_M[5]) OR ST5_A_Ca2_End) AND NOT Ins_A_Next_Cycle;

(* Section ST6_A_Rev2_左反転2: ladder, written here as Structured Text *)

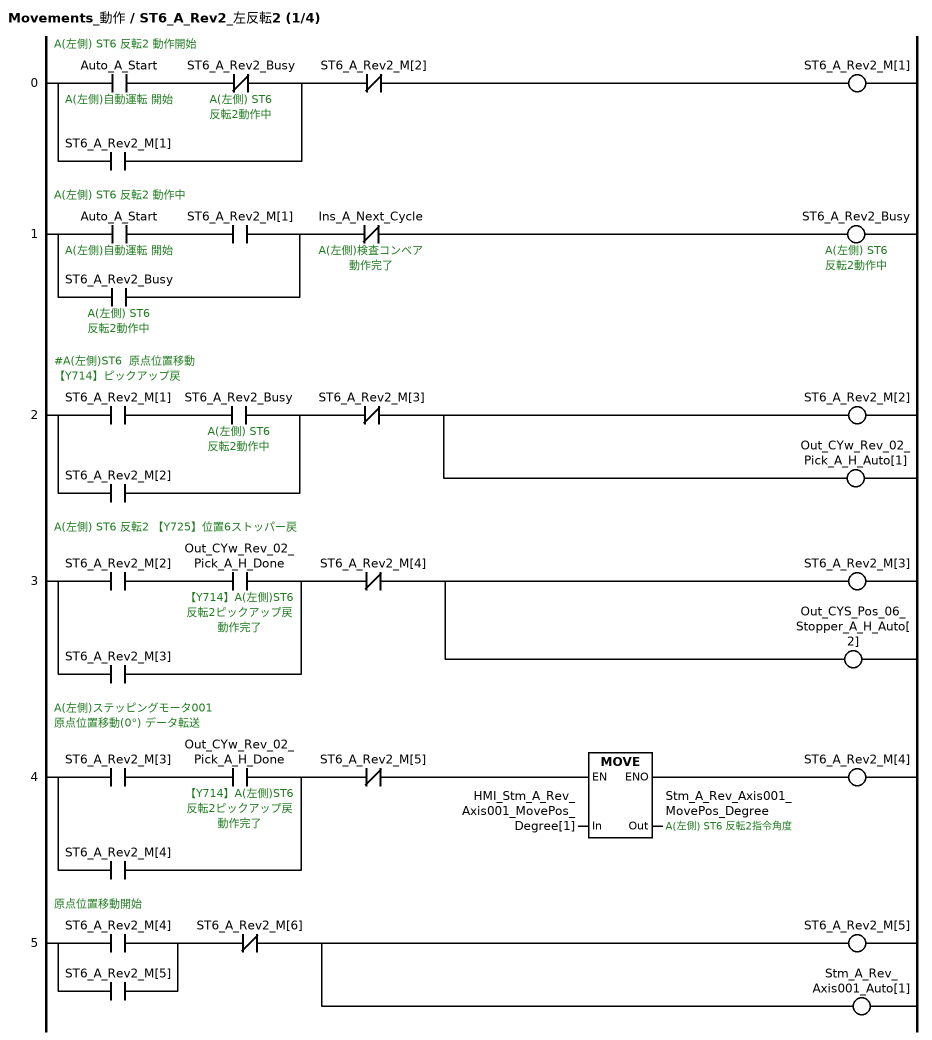
(* Rung 0: A(左側) ST6 反転2 動作開始 *)
ST6_A_Rev2_M[1] := ((Auto_A_Start AND NOT ST6_A_Rev2_Busy) OR ST6_A_Rev2_M[1]) AND NOT ST6_A_Rev2_M[2];
(* Rung 1: A(左側) ST6 反転2 動作中 *)
ST6_A_Rev2_Busy := ((Auto_A_Start AND ST6_A_Rev2_M[1]) OR ST6_A_Rev2_Busy) AND NOT Ins_A_Next_Cycle;
(* Rung 2: #A(左側)ST6  原点位置移動 / 【Y714】ピックアップ戻 *)
_p74 := ((ST6_A_Rev2_M[1] AND ST6_A_Rev2_Busy) OR ST6_A_Rev2_M[2]) AND NOT ST6_A_Rev2_M[3];
ST6_A_Rev2_M[2] := _p74;
Out_CYw_Rev_02_Pick_A_H_Auto[1] := _p74;
(* Rung 3: A(左側) ST6 反転2 【Y725】位置6ストッパー戻 *)
_p75 := ((ST6_A_Rev2_M[2] AND Out_CYw_Rev_02_Pick_A_H_Done) OR ST6_A_Rev2_M[3]) AND NOT ST6_A_Rev2_M[4];
ST6_A_Rev2_M[3] := _p75;
Out_CYS_Pos_06_Stopper_A_H_Auto[2] := _p75;
(* Rung 4: A(左側)ステッピングモータ001 / 原点位置移動(0°) データ転送 *)
IF ((ST6_A_Rev2_M[3] AND Out_CYw_Rev_02_Pick_A_H_Done) OR ST6_A_Rev2_M[4]) AND NOT ST6_A_Rev2_M[5] THEN
    Stm_A_Rev_Axis001_MovePos_Degree := HMI_Stm_A_Rev_Axis001_MovePos_Degree[1];
END_IF;
ST6_A_Rev2_M[4] := ((ST6_A_Rev2_M[3] AND Out_CYw_Rev_02_Pick_A_H_Done) OR ST6_A_Rev2_M[4]) AND NOT ST6_A_Rev2_M[5];
(* Rung 5: 原点位置移動開始 *)
_p76 := (ST6_A_Rev2_M[4] OR ST6_A_Rev2_M[5]) AND NOT ST6_A_Rev2_M[6];
ST6_A_Rev2_M[5] := _p76;
Stm_A_Rev_Axis001_Auto[1] := _p76;

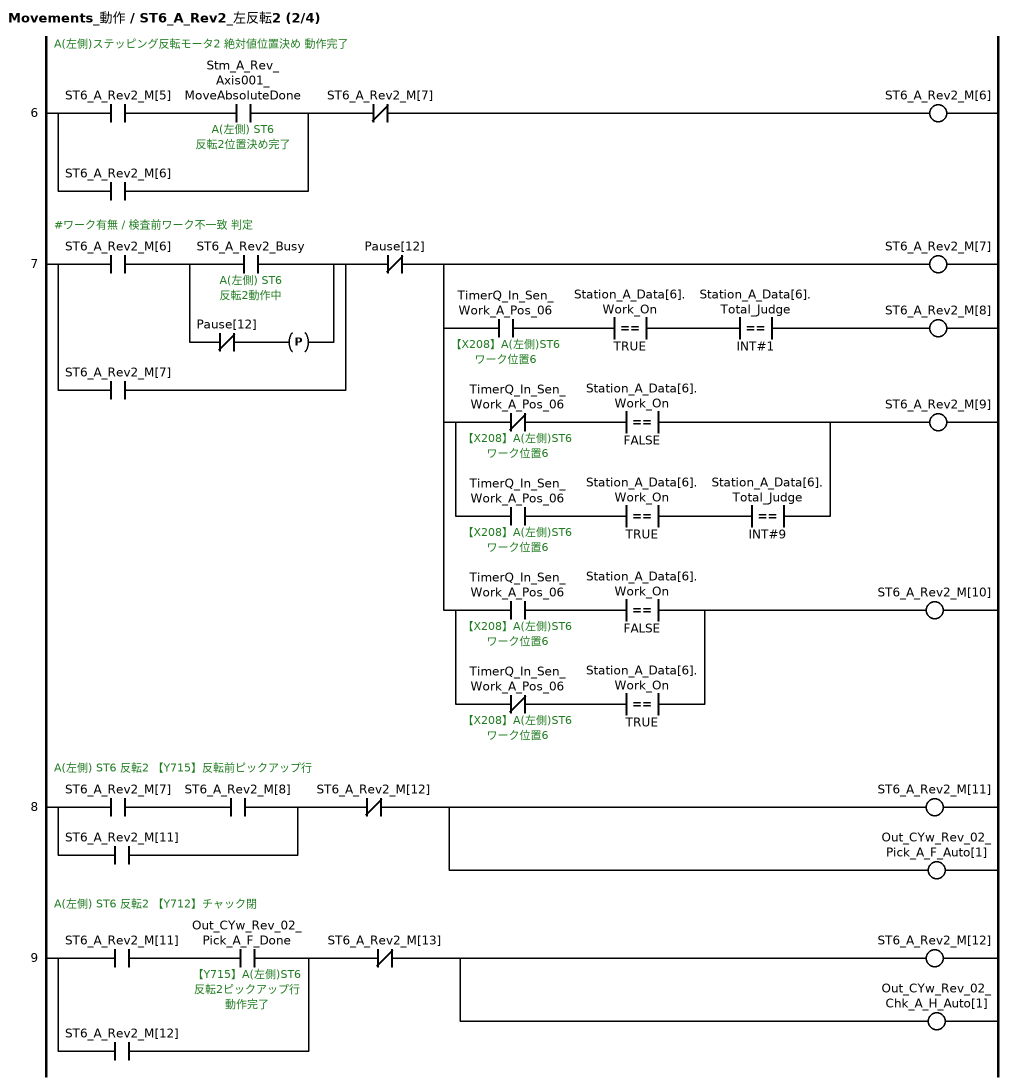
(* Rung 6: A(左側)ステッピング反転モータ2 絶対値位置決め 動作完了 *)
ST6_A_Rev2_M[6] := ((ST6_A_Rev2_M[5] AND Stm_A_Rev_Axis001_MoveAbsoluteDone) OR ST6_A_Rev2_M[6]) AND NOT ST6_A_Rev2_M[7];
(* Rung 7: #ワーク有無 / 検査前ワーク不一致 判定 *)
_e77(CLK := ST6_A_Rev2_M[6] AND NOT Pause[12]);
_p78 := ((ST6_A_Rev2_M[6] AND ST6_A_Rev2_Busy) OR _e77.Q OR ST6_A_Rev2_M[7]) AND NOT Pause[12];
ST6_A_Rev2_M[7] := _p78;
ST6_A_Rev2_M[8] := _p78 AND TimerQ_In_Sen_Work_A_Pos_06 AND (Station_A_Data[6].Work_On = TRUE) AND (Station_A_Data[6].Total_Judge = INT#1);
ST6_A_Rev2_M[9] := _p78 AND ((NOT TimerQ_In_Sen_Work_A_Pos_06 AND (Station_A_Data[6].Work_On = FALSE)) OR (TimerQ_In_Sen_Work_A_Pos_06 AND (Station_A_Data[6].Work_On = TRUE) AND (Station_A_Data[6].Total_Judge = INT#9)));
ST6_A_Rev2_M[10] := _p78 AND ((TimerQ_In_Sen_Work_A_Pos_06 AND (Station_A_Data[6].Work_On = FALSE)) OR (NOT TimerQ_In_Sen_Work_A_Pos_06 AND (Station_A_Data[6].Work_On = TRUE)));
(* Rung 8: A(左側) ST6 反転2 【Y715】反転前ピックアップ行 *)
_p79 := ((ST6_A_Rev2_M[7] AND ST6_A_Rev2_M[8]) OR ST6_A_Rev2_M[11]) AND NOT ST6_A_Rev2_M[12];
ST6_A_Rev2_M[11] := _p79;
Out_CYw_Rev_02_Pick_A_F_Auto[1] := _p79;
(* Rung 9: A(左側) ST6 反転2 【Y712】チャック閉 *)
_p80 := ((ST6_A_Rev2_M[11] AND Out_CYw_Rev_02_Pick_A_F_Done) OR ST6_A_Rev2_M[12]) AND NOT ST6_A_Rev2_M[13];
ST6_A_Rev2_M[12] := _p80;
Out_CYw_Rev_02_Chk_A_H_Auto[1] := _p80;

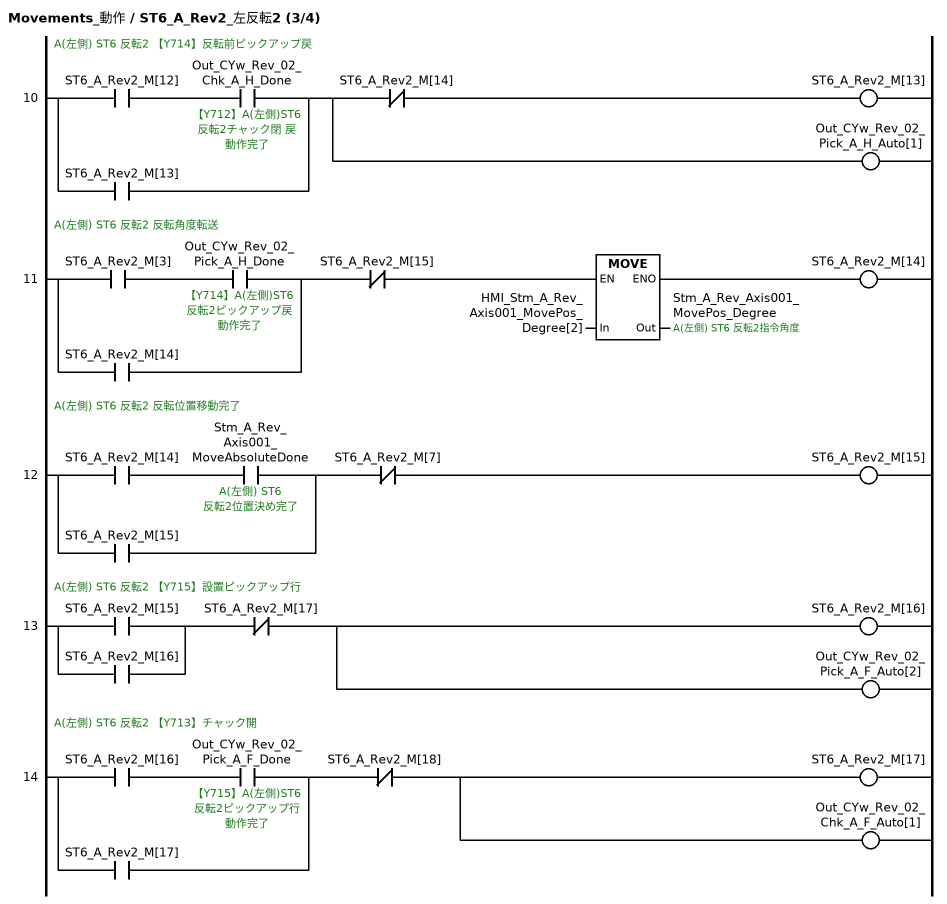
(* Rung 10: A(左側) ST6 反転2 【Y714】反転前ピックアップ戻 *)
_p81 := (ST6_A_Rev2_M[12] AND Out_CYw_Rev_02_Chk_A_H_Done) OR ST6_A_Rev2_M[13];
ST6_A_Rev2_M[13] := _p81 AND NOT ST6_A_Rev2_M[14];
Out_CYw_Rev_02_Pick_A_H_Auto[1] := _p81;
(* Rung 11: A(左側) ST6 反転2 反転角度転送 *)
IF ((ST6_A_Rev2_M[3] AND Out_CYw_Rev_02_Pick_A_H_Done) OR ST6_A_Rev2_M[14]) AND NOT ST6_A_Rev2_M[15] THEN
    Stm_A_Rev_Axis001_MovePos_Degree := HMI_Stm_A_Rev_Axis001_MovePos_Degree[2];
END_IF;
ST6_A_Rev2_M[14] := ((ST6_A_Rev2_M[3] AND Out_CYw_Rev_02_Pick_A_H_Done) OR ST6_A_Rev2_M[14]) AND NOT ST6_A_Rev2_M[15];
(* Rung 12: A(左側) ST6 反転2 反転位置移動完了 *)
ST6_A_Rev2_M[15] := ((ST6_A_Rev2_M[14] AND Stm_A_Rev_Axis001_MoveAbsoluteDone) OR ST6_A_Rev2_M[15]) AND NOT ST6_A_Rev2_M[7];
(* Rung 13: A(左側) ST6 反転2 【Y715】設置ピックアップ行 *)
_p82 := (ST6_A_Rev2_M[15] OR ST6_A_Rev2_M[16]) AND NOT ST6_A_Rev2_M[17];
ST6_A_Rev2_M[16] := _p82;
Out_CYw_Rev_02_Pick_A_F_Auto[2] := _p82;
(* Rung 14: A(左側) ST6 反転2 【Y713】チャック開 *)
_p83 := ((ST6_A_Rev2_M[16] AND Out_CYw_Rev_02_Pick_A_F_Done) OR ST6_A_Rev2_M[17]) AND NOT ST6_A_Rev2_M[18];
ST6_A_Rev2_M[17] := _p83;
Out_CYw_Rev_02_Chk_A_F_Auto[1] := _p83;

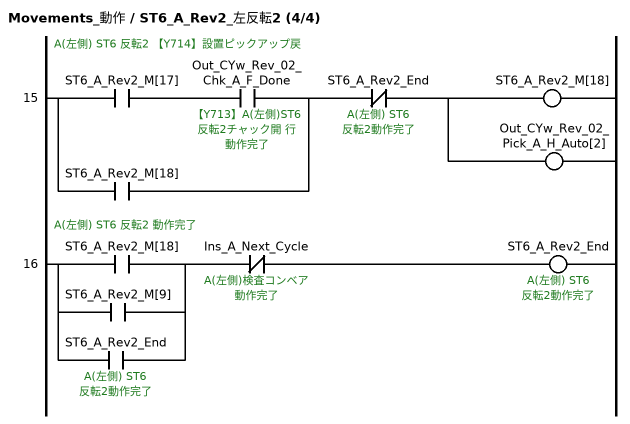
(* Rung 15: A(左側) ST6 反転2 【Y714】設置ピックアップ戻 *)
_p84 := ((ST6_A_Rev2_M[17] AND Out_CYw_Rev_02_Chk_A_F_Done) OR ST6_A_Rev2_M[18]) AND NOT ST6_A_Rev2_End;
ST6_A_Rev2_M[18] := _p84;
Out_CYw_Rev_02_Pick_A_H_Auto[2] := _p84;
(* Rung 16: A(左側) ST6 反転2 動作完了 *)
ST6_A_Rev2_End := (ST6_A_Rev2_M[18] OR ST6_A_Rev2_M[9] OR ST6_A_Rev2_End) AND NOT Ins_A_Next_Cycle;

(* Section ST7_A_Dis2_左SF排出: ladder, written here as Structured Text *)

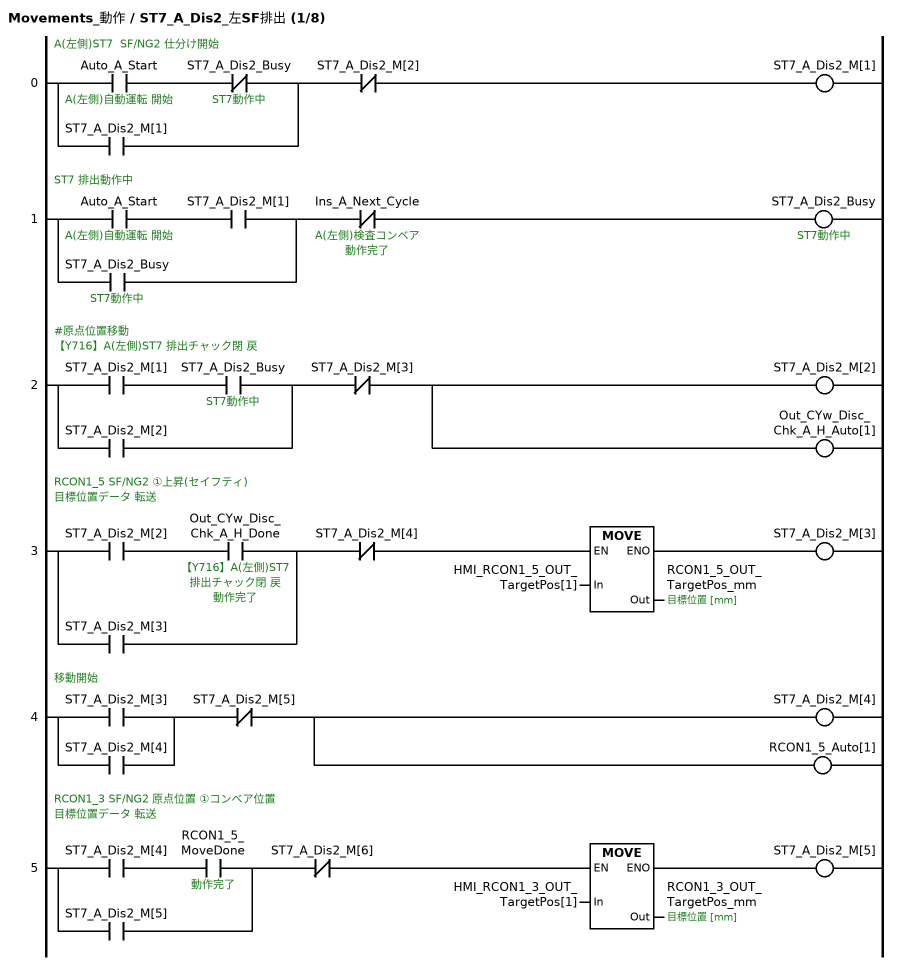
(* Rung 0: A(左側)ST7  SF/NG2 仕分け開始 *)
ST7_A_Dis2_M[1] := ((Auto_A_Start AND NOT ST7_A_Dis2_Busy) OR ST7_A_Dis2_M[1]) AND NOT ST7_A_Dis2_M[2];
(* Rung 1: ST7 排出動作中 *)
ST7_A_Dis2_Busy := ((Auto_A_Start AND ST7_A_Dis2_M[1]) OR ST7_A_Dis2_Busy) AND NOT Ins_A_Next_Cycle;
(* Rung 2: #原点位置移動 / 【Y716】A(左側)ST7 排出チャック閉 戻 *)
_p85 := ((ST7_A_Dis2_M[1] AND ST7_A_Dis2_Busy) OR ST7_A_Dis2_M[2]) AND NOT ST7_A_Dis2_M[3];
ST7_A_Dis2_M[2] := _p85;
Out_CYw_Disc_Chk_A_H_Auto[1] := _p85;
(* Rung 3: RCON1_5 SF/NG2 ①上昇(セイフティ) / 目標位置データ 転送 *)
IF ((ST7_A_Dis2_M[2] AND Out_CYw_Disc_Chk_A_H_Done) OR ST7_A_Dis2_M[3]) AND NOT ST7_A_Dis2_M[4] THEN
    RCON1_5_OUT_TargetPos_mm := HMI_RCON1_5_OUT_TargetPos[1];
END_IF;
ST7_A_Dis2_M[3] := ((ST7_A_Dis2_M[2] AND Out_CYw_Disc_Chk_A_H_Done) OR ST7_A_Dis2_M[3]) AND NOT ST7_A_Dis2_M[4];
(* Rung 4: 移動開始 *)
_p86 := (ST7_A_Dis2_M[3] OR ST7_A_Dis2_M[4]) AND NOT ST7_A_Dis2_M[5];
ST7_A_Dis2_M[4] := _p86;
RCON1_5_Auto[1] := _p86;
(* Rung 5: RCON1_3 SF/NG2 原点位置 ①コンベア位置 / 目標位置データ 転送 *)
IF ((ST7_A_Dis2_M[4] AND RCON1_5_MoveDone) OR ST7_A_Dis2_M[5]) AND NOT ST7_A_Dis2_M[6] THEN
    RCON1_3_OUT_TargetPos_mm := HMI_RCON1_3_OUT_TargetPos[1];
END_IF;
ST7_A_Dis2_M[5] := ((ST7_A_Dis2_M[4] AND RCON1_5_MoveDone) OR ST7_A_Dis2_M[5]) AND NOT ST7_A_Dis2_M[6];

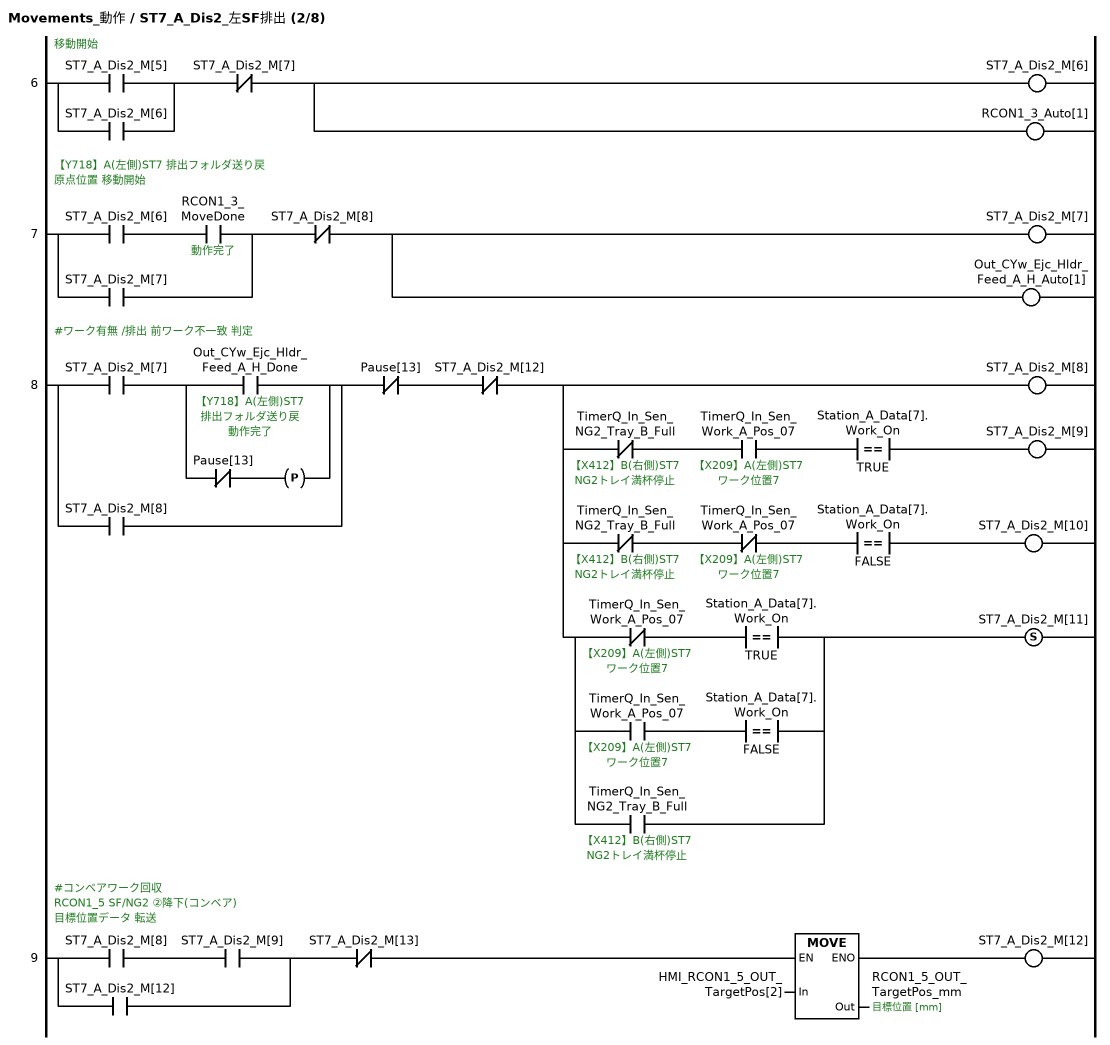
(* Rung 6: 移動開始 *)
_p87 := (ST7_A_Dis2_M[5] OR ST7_A_Dis2_M[6]) AND NOT ST7_A_Dis2_M[7];
ST7_A_Dis2_M[6] := _p87;
RCON1_3_Auto[1] := _p87;
(* Rung 7: 【Y718】A(左側)ST7 排出フォルダ送り戻 / 原点位置 移動開始 *)
_p88 := ((ST7_A_Dis2_M[6] AND RCON1_3_MoveDone) OR ST7_A_Dis2_M[7]) AND NOT ST7_A_Dis2_M[8];
ST7_A_Dis2_M[7] := _p88;
Out_CYw_Ejc_Hldr_Feed_A_H_Auto[1] := _p88;
(* Rung 8: #ワーク有無 /排出 前ワーク不一致 判定 *)
_e89(CLK := ST7_A_Dis2_M[7] AND NOT Pause[13]);
_p90 := ((ST7_A_Dis2_M[7] AND Out_CYw_Ejc_Hldr_Feed_A_H_Done) OR _e89.Q OR ST7_A_Dis2_M[8]) AND NOT Pause[13] AND NOT ST7_A_Dis2_M[12];
ST7_A_Dis2_M[8] := _p90;
ST7_A_Dis2_M[9] := _p90 AND NOT TimerQ_In_Sen_NG2_Tray_B_Full AND TimerQ_In_Sen_Work_A_Pos_07 AND (Station_A_Data[7].Work_On = TRUE);
ST7_A_Dis2_M[10] := _p90 AND NOT TimerQ_In_Sen_NG2_Tray_B_Full AND NOT TimerQ_In_Sen_Work_A_Pos_07 AND (Station_A_Data[7].Work_On = FALSE);
IF _p90 AND ((NOT TimerQ_In_Sen_Work_A_Pos_07 AND (Station_A_Data[7].Work_On = TRUE)) OR (TimerQ_In_Sen_Work_A_Pos_07 AND (Station_A_Data[7].Work_On = FALSE)) OR TimerQ_In_Sen_NG2_Tray_B_Full) THEN
    ST7_A_Dis2_M[11] := TRUE;
END_IF;
(* Rung 9: #コンベアワーク回収 / RCON1_5 SF/NG2 ②降下(コンベア) / 目標位置データ 転送 *)
IF ((ST7_A_Dis2_M[8] AND ST7_A_Dis2_M[9]) OR ST7_A_Dis2_M[12]) AND NOT ST7_A_Dis2_M[13] THEN
    RCON1_5_OUT_TargetPos_mm := HMI_RCON1_5_OUT_TargetPos[2];
END_IF;
ST7_A_Dis2_M[12] := ((ST7_A_Dis2_M[8] AND ST7_A_Dis2_M[9]) OR ST7_A_Dis2_M[12]) AND NOT ST7_A_Dis2_M[13];

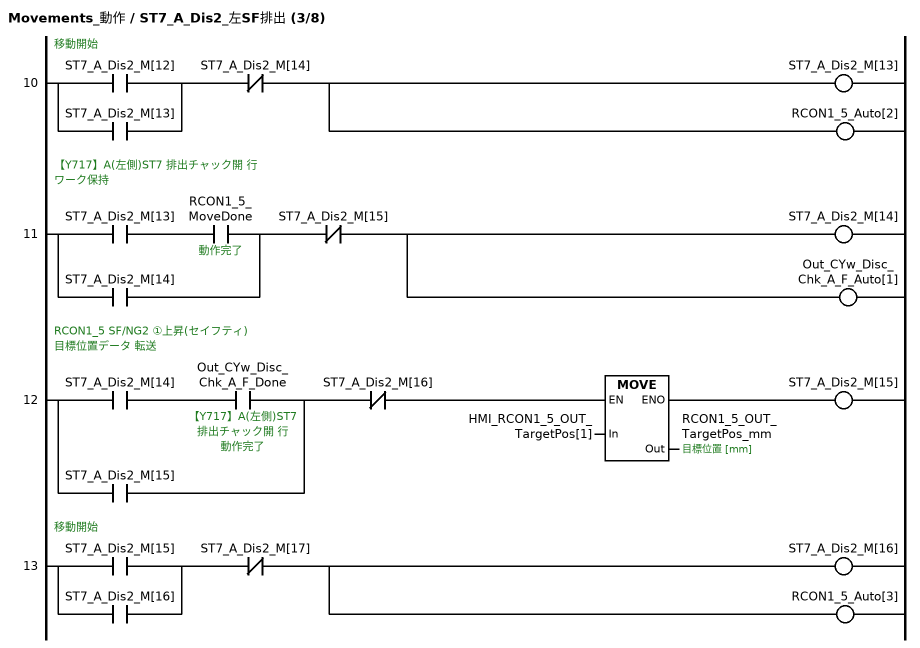
(* Rung 10: 移動開始 *)
_p91 := (ST7_A_Dis2_M[12] OR ST7_A_Dis2_M[13]) AND NOT ST7_A_Dis2_M[14];
ST7_A_Dis2_M[13] := _p91;
RCON1_5_Auto[2] := _p91;
(* Rung 11: 【Y717】A(左側)ST7 排出チャック開 行 / ワーク保持 *)
_p92 := ((ST7_A_Dis2_M[13] AND RCON1_5_MoveDone) OR ST7_A_Dis2_M[14]) AND NOT ST7_A_Dis2_M[15];
ST7_A_Dis2_M[14] := _p92;
Out_CYw_Disc_Chk_A_F_Auto[1] := _p92;
(* Rung 12: RCON1_5 SF/NG2 ①上昇(セイフティ) / 目標位置データ 転送 *)
IF ((ST7_A_Dis2_M[14] AND Out_CYw_Disc_Chk_A_F_Done) OR ST7_A_Dis2_M[15]) AND NOT ST7_A_Dis2_M[16] THEN
    RCON1_5_OUT_TargetPos_mm := HMI_RCON1_5_OUT_TargetPos[1];
END_IF;
ST7_A_Dis2_M[15] := ((ST7_A_Dis2_M[14] AND Out_CYw_Disc_Chk_A_F_Done) OR ST7_A_Dis2_M[15]) AND NOT ST7_A_Dis2_M[16];
(* Rung 13: 移動開始 *)
_p93 := (ST7_A_Dis2_M[15] OR ST7_A_Dis2_M[16]) AND NOT ST7_A_Dis2_M[17];
ST7_A_Dis2_M[16] := _p93;
RCON1_5_Auto[3] := _p93;

